(* IEC 61131-3 sources: Industry-PLC-LLM/data/PLCBEAD_repo/PLCBEAD_PLCEmbed-main/PLC-BEAD/Source/PLC_Programs (part 12) *)

(* ---- TEMP_EXT.ST ---- *)
FUNCTION UDINT_TO_TIME2:TIME

	VAR_INPUT
		IN :	UDINT;
	END_VAR

	UDINT_TO_TIME2 := DINT_TO_TIME(UDINT_TO_DINT(IN));

END_FUNCTION

FUNCTION_BLOCK T_PLC_MS_block
	VAR_OUTPUT
		T_PLC_MS :	UDINT;
	END_VAR

	VAR_EXTERNAL
		PLC_TICKS_PER_SEC :	INT;
		PLC_SYS_TICK_CNT :	DINT;
	END_VAR

	VAR
		debug :	BOOL;(*Debug-Mode ON / OFF*)
		N :	INT;(*Debug-Faktor*)
		Offset :	UDINT;(*Debug-Offset*)
		temp :	DWORD := DWORD#1;(*Debug-Offset*)
		mode :	BOOL;(*modus*)
		faktor :	UDINT;(*Systemtakt-Faktor*)
		init :	BOOL;
		v_plc_ticks_per_sec :	UDINT;
		base :	UDINT := UDINT#1000;
	END_VAR

	IF init = FALSE THEN
		v_plc_ticks_per_sec := INT_TO_UDINT(PLC_TICKS_PER_SEC);
		IF v_plc_ticks_per_sec = UDINT#1024 THEN
			faktor := UDINT#1;
			mode := FALSE;
		ELSIF v_plc_ticks_per_sec > UDINT#0 THEN
			IF v_plc_ticks_per_sec <= base THEN
				faktor := base / v_plc_ticks_per_sec;
				mode := FALSE;
			ELSE
				faktor := v_plc_ticks_per_sec / base;
				mode := TRUE;
			END_IF;
		ELSE
			faktor := UDINT#1;
		END_IF;
		init := TRUE;
	END_IF;

	IF mode THEN
		T_PLC_MS := DINT_TO_UDINT(PLC_SYS_TICK_CNT) / faktor;
	ELSE
		T_PLC_MS := DINT_TO_UDINT(PLC_SYS_TICK_CNT) * faktor;
	END_IF;

	IF debug THEN
		T_PLC_MS := (DWORD_TO_UDINT(SHL(UDINT_TO_DWORD(T_PLC_MS),N) OR SHL(temp,N)) - UDINT#1) + Offset;
	END_IF;
END_FUNCTION_BLOCK

FUNCTION _INT_TO_UDINT:UDINT
	VAR_INPUT
		IN :	INT;
	END_VAR

	_INT_TO_UDINT := DINT_TO_UDINT(INT_TO_DINT(IN));
END_FUNCTION

FUNCTION SET_DATE:UDINT

	VAR_INPUT
		YEAR :	INT;
		MONTH :	INT;
		DAY :	INT;
	END_VAR

	VAR
		count :	INT;
	END_VAR

	IF month > 2 THEN
		count := (month - 1) * 30;
		IF month > 7 THEN
			count := count + DWORD_TO_INT(SHR(DINT_TO_DWORD(INT_TO_DINT(month) - INT_TO_DINT(3)),1));
		ELSE
			count := count + DWORD_TO_INT(SHR(DINT_TO_DWORD(INT_TO_DINT(month) - INT_TO_DINT(4)),1));
		END_IF;
		IF SHL(INT_TO_WORD(year),14) = WORD#0 THEN
			count := count + 1;
		END_IF;
	ELSE
		count := (month - 1) * 31;
	END_IF;
	SET_DATE := (_INT_TO_UDINT(count + day - 1) + DWORD_TO_UDINT(SHR(UDINT_TO_DWORD(_INT_TO_UDINT(year) * UDINT#1461 - UDINT#2878169), 2))) * UDINT#86400;

END_FUNCTION

FUNCTION LEAP_OF_DATE:BOOL

	VAR_INPUT
		IDATE :	UDINT;
	END_VAR

	LEAP_OF_DATE := SHL(UDINT_TO_DWORD((idate + UDINT#43200) / UDINT#31557600), 30) = DWORD#16#80000000;

END_FUNCTION

FUNCTION DAY_OF_YEAR:INT
	VAR_INPUT
		IDATE :	DATE;
	END_VAR

	DAY_OF_YEAR := UDINT_TO_INT((DATE_TO_UDINT(idate) / UDINT#86400) MOD UDINT#1461);
	IF DAY_OF_YEAR > 729 THEN
		IF DAY_OF_YEAR > 1095 THEN DAY_OF_YEAR := DAY_OF_YEAR - 1095; ELSE DAY_OF_YEAR := DAY_OF_YEAR - 729; END_IF;
	ELSIF DAY_OF_YEAR > 364 THEN
		DAY_OF_YEAR := DAY_OF_YEAR - 364;
	ELSE
		DAY_OF_YEAR := DAY_OF_YEAR + 1;
	END_IF;
END_FUNCTION

FUNCTION DAY_OF_YEAR_UDINT:INT
	VAR_INPUT
		IDATE :	UDINT;
	END_VAR

	DAY_OF_YEAR_UDINT := UDINT_TO_INT((idate / UDINT#86400) MOD UDINT#1461);
	IF DAY_OF_YEAR_UDINT > 729 THEN
		IF DAY_OF_YEAR_UDINT > 1095 THEN DAY_OF_YEAR_UDINT := DAY_OF_YEAR_UDINT - 1095; ELSE DAY_OF_YEAR_UDINT := DAY_OF_YEAR_UDINT - 729; END_IF;
	ELSIF DAY_OF_YEAR_UDINT > 364 THEN
		DAY_OF_YEAR_UDINT := DAY_OF_YEAR_UDINT - 364;
	ELSE
		DAY_OF_YEAR_UDINT := DAY_OF_YEAR_UDINT + 1;
	END_IF;
END_FUNCTION

FUNCTION MONTH_OF_DATE_UDINT:INT

	VAR_INPUT
		IDATE :	UDINT;
	END_VAR

	MONTH_OF_DATE_UDINT := DAY_OF_YEAR_UDINT(idate);
	IF MONTH_OF_DATE_UDINT < 32 THEN
		MONTH_OF_DATE_UDINT := 1;
	ELSIF LEAP_OF_DATE(IDATE) THEN
		MONTH_OF_DATE_UDINT := (MONTH_OF_DATE_UDINT * 53 + 1668) / 1623;
	ELSE
		MONTH_OF_DATE_UDINT := (MONTH_OF_DATE_UDINT * 53 + 1700) / 1620;
	END_IF;

END_FUNCTION

FUNCTION DAY_OF_MONTH:INT
	VAR_INPUT
		IDATE :	UDINT;
	END_VAR

	day_of_month := day_of_year_UDINT(idate);

	IF leap_of_Date(idate) THEN
		CASE day_of_month OF
			32..60	:	day_of_month := day_of_month - 31;
			61..91	:	day_of_month := day_of_month - 60;
			92..121 :	day_of_month := day_of_month - 91;
			122..152:	day_of_month := day_of_month - 121;
			153..182:	day_of_month := day_of_month - 152;
			183..213:	day_of_month := day_of_month - 182;
			214..244:	day_of_month := day_of_month - 213;
			245..274:	day_of_month := day_of_month - 244;
			275..305:	day_of_month := day_of_month - 274;
			306..335:	day_of_month := day_of_month - 305;
			336..366:	day_of_month := day_of_month - 335;
		END_CASE;
	ELSE
		CASE day_of_month OF
			32..59	:	day_of_month := day_of_month - 31;
			60..90	:	day_of_month := day_of_month - 59;
			91..120 :	day_of_month := day_of_month - 90;
			121..151:	day_of_month := day_of_month - 120;
			152..181:	day_of_month := day_of_month - 151;
			182..212:	day_of_month := day_of_month - 181;
			213..243:	day_of_month := day_of_month - 212;
			244..273:	day_of_month := day_of_month - 243;
			274..304:	day_of_month := day_of_month - 273;
			305..334:	day_of_month := day_of_month - 304;
			335..365:	day_of_month := day_of_month - 334;
		END_CASE;
	END_IF;

END_FUNCTION

FUNCTION MID3:REAL

	VAR_INPUT
		IN1 :	REAL;
		IN2 :	REAL;
		IN3 :	REAL;
	END_VAR

	VAR
		_IN1 :	REAL;
		_IN2 :	REAL;
		_IN3 :	REAL;
	END_VAR

	_IN1 := IN1;
	_IN2 := IN2;
	_IN3 := IN3;

	IF _IN1 > _IN2 THEN MID3 := _IN1; _IN1 := _IN2; _IN2 := MID3; END_IF;
	IF _IN2 > _IN3 THEN _IN2 := _IN3; END_IF;
	MID3 := SEL(_IN1 > _IN2, _IN2, _IN1);

END_FUNCTION

FUNCTION _BYTE_TO_INT:INT
	VAR_INPUT
		IN :	BYTE;
	END_VAR

	_BYTE_TO_INT := USINT_TO_INT(BYTE_TO_USINT(IN));
END_FUNCTION

FUNCTION MULTI_IN:REAL

	VAR_INPUT
		IN_1 :	REAL;
		IN_2 :	REAL;
		IN_3 :	REAL;
		DEFAULT :	REAL;
		IN_MIN :	REAL;
		IN_MAX :	REAL;
		MODE :	BYTE;
	END_VAR

	VAR
		count :	INT;
		F1 :	BOOL;
		F2 :	BOOL;
		F3 :	BOOL;
	END_VAR

	F1 :=  in_1 > in_min AND in_1 < in_max;
	F2 :=  in_2 > in_min AND in_2 < in_max;
	F3 :=  in_3 > in_min AND in_3 < in_max;

	CASE _BYTE_TO_INT(mode) OF
	0:	count := 0;
		IF F1 THEN
			count := count + 1;
			MULTI_IN := in_1;
		ELSE
			MULTI_IN := 0.0;
		END_IF;
		IF F2 THEN
			count := count + 1;
			MULTI_IN := MULTI_IN + in_2;
		END_IF;
		IF F3 THEN
			count := count + 1;
			MULTI_IN := MULTI_IN + in_3;
		END_IF;
		MULTI_IN := SEL_REAL(count = 0, MULTI_IN / INT_TO_REAL(count), default);

	1:	MULTI_IN := SEL_REAL(F1, default, IN_1);

	2:	MULTI_IN := SEL_REAL(F2, default, IN_2);

	3:	MULTI_IN := SEL_REAL(F3, default, IN_3);

	4:	MULTI_IN := default;

	5:	MULTI_IN := SEL_REAL(F1, in_max, IN_1);
		IF F2 AND in_2 < MULTI_IN THEN MULTI_IN := in_2; END_IF;
		IF F3 AND in_3 < MULTI_IN THEN MULTI_IN := in_3; END_IF;
		IF MULTI_IN = in_max THEN MULTI_IN := default; END_IF;

	6:	MULTI_IN := SEL_REAL(F1, in_min, IN_1);
		IF F2 AND in_2 > MULTI_IN THEN MULTI_IN := in_2; END_IF;
		IF F3 AND in_3 > MULTI_IN THEN MULTI_IN := in_3; END_IF;
		IF MULTI_IN = in_min THEN MULTI_IN := default; END_IF;

	7:	IF F1 AND F2 AND F3 THEN MULTI_IN := MID3(in_1, in_2, in_3);
		ELSIF F1 AND F2 THEN MULTI_IN := MIN(in_1, in_2);
		ELSIF F1 AND F3 THEN MULTI_IN := MIN(in_1, in_3);
		ELSIF F2 AND F3 THEN MULTI_IN := MIN(in_2, in_3);
		ELSIF F1 THEN MULTI_IN := in_1;
		ELSIF F2 THEN MULTI_IN := in_2;
		ELSIF F3 THEN MULTI_IN := in_3;
		ELSE MULTI_IN := default;
		END_IF;

	END_CASE;

END_FUNCTION

FUNCTION _DT_TO_DATE_B:UDINT

	VAR_INPUT
		_INN :	UDINT;
	END_VAR

	_DT_TO_DATE_B := (_INN / UDINT#86400) * UDINT#86400;
END_FUNCTION

FUNCTION DT_TO_TOD2:UDINT
	VAR_INPUT
		IN :	UDINT;
	END_VAR

	DT_TO_TOD2 := (IN MOD UDINT#86400) * UDINT#1000;
END_FUNCTION

FUNCTION_BLOCK TEMP_EXT_Block

	VAR_INPUT
		T_EXT1 :	REAL;
		T_EXT2 :	REAL;
		T_EXT3 :	REAL;
		T_EXT_CONFIG :	BYTE := 0;
		DT_IN :	UDINT;
		T_EXT_MIN :	REAL := REAL#-40.0;
		T_EXT_MAX :	REAL := REAL#60.0;
		T_EXT_DEFAULT :	REAL := REAL#-10.0;
		HEAT_PERIOD_START :	UDINT := UDINT#20995200;
		HEAT_PERIOD_STOP :	UDINT := UDINT#10281600;
		COOL_PERIOD_START :	UDINT := UDINT#07776000;
		COOL_PERIOD_STOP :	UDINT := UDINT#23500800;
		HEAT_START_TEMP_DAY :	REAL := REAL#15.0;
		HEAT_START_TEMP_NIGHT :	REAL := REAL#10.0;
		HEAT_STOP_TEMP :	REAL := REAL#18.0;
		COOL_START_TEMP_DAY :	REAL := REAL#26.0;
		COOL_START_TEMP_NIGHT :	REAL := REAL#26.0;
		COOL_STOP_TEMP :	REAL := REAL#24.0;
		START_DAY :	UDINT := UDINT#32400000;
		START_NIGHT :	UDINT := UDINT#75600000;
		CYCLE_TIME :	TIME := t#10m;
	END_VAR

	VAR_OUTPUT
		T_EXT :	REAL;
		HEAT :	BOOL;
		COOL :	BOOL;
	END_VAR

	VAR
		tx :	TIME;
		last_run :	TIME;
		init :	BOOL;
		cool_start :	UDINT;
		cool_stop :	UDINT;
		heat_start :	UDINT;
		heat_stop :	UDINT;
		xdate :	UDINT;
		day :	BOOL;
		T_PLC_MS :	T_PLC_MS_Block;
	END_VAR

	IF NOT init THEN
		init := TRUE;
		heat_start := SET_DATE(1972,MONTH_OF_DATE_UDINT(heat_period_start),DAY_OF_MONTH(heat_period_start));
		heat_stop := SET_DATE(1972,MONTH_OF_DATE_UDINT(heat_period_stop),DAY_OF_MONTH(heat_period_stop));
		cool_start := SET_DATE(1972,MONTH_OF_DATE_UDINT(cool_period_start),DAY_OF_MONTH(cool_period_start));
		cool_stop := SET_DATE(1972,MONTH_OF_DATE_UDINT(cool_period_stop),DAY_OF_MONTH(cool_period_stop));
	END_IF;

	T_PLC_MS();
	tx:= UDINT_TO_TIME(T_PLC_MS.T_PLC_MS);

	IF tx - last_run < cycle_time THEN RETURN; END_IF;

	xdate := SET_DATE(1972,MONTH_OF_DATE_UDINT(_DT_TO_DATE_B(dt_in)),DAY_OF_MONTH(_DT_TO_DATE_B(dt_in)));
	day := DT_TO_TOD2(dt_in) >= start_day AND  DT_TO_TOD2(dt_in) < start_night;

	t_ext := MULTI_IN(t_ext1, t_ext2, t_ext3, t_ext_default, t_ext_min, t_ext_max, t_ext_config);

	IF (heat_start <= heat_stop AND xdate >= heat_start AND xdate <= heat_stop) OR (heat_start > heat_stop AND (xdate >= heat_start OR xdate <= heat_stop)) THEN
		IF day AND t_ext <= heat_start_temp_day THEN
			heat := TRUE;
		ELSIF NOT day AND t_ext <= heat_start_temp_night THEN
			heat := TRUE;
		ELSIF t_ext >= heat_stop_temp THEN
			heat := FALSE;
		END_IF;
	ELSE
		heat := FALSE;
	END_IF;

	IF (cool_start <= cool_stop AND xdate >= cool_start AND xdate <= cool_stop) OR (cool_start > cool_stop AND (xdate >= cool_start OR xdate <= cool_stop)) THEN
		IF day AND t_ext >= cool_start_temp_day THEN
			cool := TRUE;
		ELSIF NOT day AND t_ext >= cool_start_temp_night THEN
			cool := TRUE;
		ELSIF t_ext <= cool_stop_temp THEN
			cool := FALSE;
		END_IF;
	ELSE
		cool := FALSE;
	END_IF;

	last_run := tx;

END_FUNCTION_BLOCK

PROGRAM program0
	VAR
		T_EXT1 :	REAL;
		T_EXT2 :	REAL;
		T_EXT3 :	REAL;
		T_EXT_CONFIG :	BYTE := 0;
		DT_IN :	UDINT;
		T_EXT_MIN :	REAL := REAL#-40.0;
		T_EXT_MAX :	REAL := REAL#60.0;
		T_EXT_DEFAULT :	REAL := REAL#-10.0;
		HEAT_PERIOD_START :	UDINT := UDINT#20995200;
		HEAT_PERIOD_STOP :	UDINT := UDINT#10281600;
		COOL_PERIOD_START :	UDINT := UDINT#07776000;
		COOL_PERIOD_STOP :	UDINT := UDINT#23500800;
		HEAT_START_TEMP_DAY :	REAL := REAL#15.0;
		HEAT_START_TEMP_NIGHT :	REAL := REAL#10.0;
		HEAT_STOP_TEMP :	REAL := REAL#18.0;
		COOL_START_TEMP_DAY :	REAL := REAL#26.0;
		COOL_START_TEMP_NIGHT :	REAL := REAL#26.0;
		COOL_STOP_TEMP :	REAL := REAL#24.0;
		START_DAY :	UDINT := UDINT#32400000;
		START_NIGHT :	UDINT := UDINT#75600000;
		CYCLE_TIME :	TIME := t#10m;
		T_EXT :	REAL;
		HEAT :	BOOL;
		COOL :	BOOL;

		func_block : TEMP_EXT_Block;
	END_VAR

	func_block.T_EXT1 := T_EXT1;
	func_block.T_EXT2 := T_EXT2;
	func_block.T_EXT3 := T_EXT3 ;
	func_block.T_EXT_CONFIG := T_EXT_CONFIG;
	func_block.DT_IN := DT_IN;
	func_block.T_EXT_MIN := T_EXT_MIN ;
	func_block.T_EXT_MAX := T_EXT_MAX;
	func_block.T_EXT_DEFAULT := T_EXT_DEFAULT;
	func_block.HEAT_PERIOD_START := HEAT_PERIOD_START ;
	func_block.HEAT_PERIOD_STOP := HEAT_PERIOD_STOP;
	func_block.COOL_PERIOD_START := COOL_PERIOD_START;
	func_block.COOL_PERIOD_STOP := COOL_PERIOD_STOP ;
	func_block.HEAT_START_TEMP_DAY := HEAT_START_TEMP_DAY;
	func_block.HEAT_START_TEMP_NIGHT := HEAT_START_TEMP_NIGHT;
	func_block.HEAT_STOP_TEMP := HEAT_STOP_TEMP ;
	func_block.COOL_START_TEMP_DAY := COOL_START_TEMP_DAY;
	func_block.COOL_START_TEMP_NIGHT := COOL_START_TEMP_NIGHT;
	func_block.COOL_STOP_TEMP:= COOL_STOP_TEMP ;
	func_block.START_DAY := START_DAY;
	func_block.START_NIGHT := START_NIGHT;
	func_block.CYCLE_TIME:= CYCLE_TIME ;

	func_block();
	T_EXT  := func_block.T_EXT;
	HEAT  := func_block.HEAT;
	COOL  := func_block.COOL;

END_PROGRAM

CONFIGURATION Config0
	VAR_GLOBAL
		PLC_TICKS_PER_SEC :	INT;
		PLC_SYS_TICK_CNT :	DINT;
	END_VAR
  	RESOURCE Res0 ON PLC
    	TASK task0(INTERVAL := T#20ms,PRIORITY := 0);
    	PROGRAM instance0 WITH task0 : program0;
  	END_RESOURCE
END_CONFIGURATION

(* ---- TEMPERATURE.ST ---- *)
FUNCTION_BLOCK TEMPERATURE

	VAR_INPUT
		K :	REAL;
		C :	REAL := -273.15;
		F :	REAL := -459.67;
		RE :	REAL := -218.52;
		RA :	REAL := 0.0;
	END_VAR

	VAR_OUTPUT
		YK :	REAL;
		YC :	REAL;
		YF :	REAL;
		YRE :	REAL;
		YRA :	REAL;
	END_VAR

	YK := K + (C + 273.15) + (F + 459.67) * 0.555555555555 + (Re * 1.25 + 273.15) + (Ra * 0.555555555555);
	YC := YK -273.15;
	YF := YK * 1.8 - 459.67;
	YRe := (YK - 273.15) * 0.8;
	YRa := YK * 1.8;

END_FUNCTION_BLOCK

PROGRAM program0
  VAR
	K :	REAL;
	C :	REAL := -273.15;
	F :	REAL := -459.67;
	RE :	REAL := -218.52;
	RA :	REAL := 0.0;
	YK :	REAL;
	YC :	REAL;
	YF :	REAL;
	YRE :	REAL;
	YRA :	REAL;
	func_block : TEMPERATURE;
  END_VAR
	func_block.K  :=K;
	func_block.C  :=C;
	func_block.F  :=F;
	func_block.RE  :=RE;
	func_block.RA  :=RA;
	func_block();
	YK := func_block.YK;
	YC := func_block.YC;
	YF := func_block.YF;
	YRE := func_block.YRE;
	YRA := func_block.YRA;

END_PROGRAM

CONFIGURATION Config0
	RESOURCE Res0 ON PLC
		TASK task0(INTERVAL := T#20ms,PRIORITY := 0);
		PROGRAM instance0 WITH task0 : program0;
	END_RESOURCE
END_CONFIGURATION

(* ---- TICKER.ST ---- *)
TYPE
	oscat_delay_buf             : ARRAY [0..31]   OF REAL;
END_TYPE

FUNCTION INC1:INT

	VAR_INPUT
		X :	INT;
		N :	INT;
	END_VAR

	IF X >= N - 1 THEN
		INC1 := 0;
	ELSE
		INC1 := X + 1;
	END_IF;
END_FUNCTION

FUNCTION_BLOCK DELAY

	VAR_INPUT
		IN :	REAL;
		N :	INT;
		RST :	BOOL;
	END_VAR

	VAR_OUTPUT
		OUT :	REAL;
	END_VAR

	VAR
		buf :	oscat_delay_buf;
		i :	INT;
		init :	BOOL;
		stop :	INT;
	END_VAR

	stop := LIMIT(0,N,32) - 1;
	IF rst OR NOT init THEN
		init := TRUE;
		FOR i := 0 TO stop DO buf[i] := in; END_FOR;
		out := in;
		i := 0;
	ELSIF stop < 0 THEN
		out := in;
	ELSE
		out := buf[i];
		buf[i] := in;
		i := INC1(i, N);
	END_IF;

END_FUNCTION_BLOCK

FUNCTION_BLOCK TICKER

	VAR_INPUT
		N :	INT;
		PT :	TIME;
		TEXT :	STRING;
	END_VAR

	VAR_OUTPUT
		DISPLAY :	STRING;
	END_VAR

	VAR
		_delay :	TP;
		rollout :	STRING;
		text_len :	INT;
		rollout_step :	INT;
		_step :	INT;
	END_VAR

	text_len := LEN(text);

	IF N < text_len THEN
		IF NOT _delay.Q THEN

			IF _step > text_len THEN
				rollout_step := 0;
				rollout := '';
				_step := 0;
			END_IF;

			IF _step + N > text_len THEN
				_step := _step + 1;
				rollout_step := rollout_step +1;
				display := MID(text, N - rollout_step, _step);
				rollout := CONCAT(rollout,'#');
				display := CONCAT(display,rollout);
			ELSE
				_step := _step + 1;
				display := MID(text, N, _step);
			END_IF;
			_delay(TRUE, PT);
		ELSE
			_delay(FALSE);
		END_IF;
	ELSE
		display := text;
	END_IF;

END_FUNCTION_BLOCK

PROGRAM program0
	VAR
		N :	INT;
		PT :	TIME;
		TEXT :	STRING;
		DISPLAY :	STRING;
		func_block : TICKER;
  	END_VAR
	func_block.N  :=N;
	func_block.PT  :=PT;
	func_block.TEXT  :=TEXT;
	func_block();
	DISPLAY := func_block.DISPLAY;
END_PROGRAM

CONFIGURATION Config0
	RESOURCE Res0 ON PLC
		TASK task0(INTERVAL := T#20ms,PRIORITY := 0);
		PROGRAM instance0 WITH task0 : program0;
	END_RESOURCE
END_CONFIGURATION

(* ---- TIMER_1.ST ---- *)
FUNCTION TIMECHECK:BOOL

	VAR_INPUT
		TD :	UDINT;
		START :	UDINT;
		STOP :	UDINT;
	END_VAR

	IF stop < start THEN
		TIMECHECK := start <= TD OR  TD < stop;
	ELSE
		TIMECHECK := start <= TD AND TD < stop;
	END_IF;

END_FUNCTION

FUNCTION TIME_TO_TOD:UDINT

	VAR_INPUT
		IN :	TIME;
	END_VAR

	TIME_TO_TOD := DWORD_TO_UDINT(TIME_TO_DWORD(IN));
END_FUNCTION

FUNCTION TOD_TO_TIME:TIME
	VAR_INPUT
		IN :	UDINT;
	END_VAR

	TOD_TO_TIME := DWORD_TO_TIME(UDINT_TO_DWORD(IN));
END_FUNCTION

FUNCTION DAY_OF_WEEK:INT
  VAR_INPUT
    IDATE :	UDINT;
  END_VAR

  DAY_OF_WEEK := UDINT_TO_INT((idate / UDINT#86400 + UDINT#3) MOD UDINT#7) + INT#01;
END_FUNCTION

FUNCTION _DT_TO_DATE_B:UDINT

	VAR_INPUT
		_INN :	UDINT;
	END_VAR

	_DT_TO_DATE_B := (_INN / UDINT#86400) * UDINT#86400;
END_FUNCTION

FUNCTION DT_TO_TOD2:UDINT
	VAR_INPUT
		IN :	UDINT;
	END_VAR

	DT_TO_TOD2 := (IN MOD UDINT#86400) * UDINT#1000;
END_FUNCTION

FUNCTION TIME_TO_TOD2:UDINT

	VAR_INPUT
		IN :	TIME;
	END_VAR

	TIME_TO_TOD2 := DWORD_TO_UDINT(TIME_TO_DWORD(IN));
END_FUNCTION

FUNCTION_BLOCK TIMER_1_Block

	VAR_INPUT
		E :	BOOL := TRUE;
		DTI :	UDINT;
		START :	UDINT;
		DURATION :	TIME;
		DAY :	BYTE := BYTE#2#0111_1111;
	END_VAR

	VAR_OUTPUT
		Q :	BOOL;
		STOP :	TIME;
	END_VAR

	IF E THEN
		stop := TOD_TO_TIME(START) + DURATION;
		IF stop > T#24h THEN stop := stop - T#24h; END_IF;
		Q := TIMECHECK(DT_TO_TOD2(DTI), START, TIME_TO_TOD2(stop)) AND (SHR(BYTE#128, DAY_OF_WEEK(_DT_TO_DATE_B(DTI))) AND DAY) > BYTE#0;
	ELSE
		Q := FALSE;
	END_IF;

END_FUNCTION_BLOCK

PROGRAM program0
	VAR
		E :	BOOL := TRUE;
		DTI :	UDINT;
		START :	UDINT;
		DURATION :	TIME;
		DAY :	BYTE := BYTE#2#0111_1111;
		Q :	BOOL;
		STOP :	TIME;

		func_block : TIMER_1_Block;
	END_VAR
	func_block.E := E;
	func_block.DTI := DTI;
	func_block.START := START ;
	func_block.DURATION    := DURATION    ;
	func_block.DAY := DAY;

	func_block();
	Q  := func_block.Q;
	STOP  := func_block.STOP;
END_PROGRAM

CONFIGURATION Config0
	RESOURCE Res0 ON PLC
		TASK task0(INTERVAL := T#20ms,PRIORITY := 0);
		PROGRAM instance0 WITH task0 : program0;
	END_RESOURCE
END_CONFIGURATION

(* ---- TIMER_2.ST ---- *)
FUNCTION UDINT_TO_TIME2:TIME

	VAR_INPUT
		IN :	UDINT;
	END_VAR

	UDINT_TO_TIME2 := DINT_TO_TIME(UDINT_TO_DINT(IN));

END_FUNCTION

FUNCTION_BLOCK T_PLC_MS_block
	VAR_OUTPUT
		T_PLC_MS :	UDINT;
	END_VAR

	VAR_EXTERNAL
		PLC_TICKS_PER_SEC :	INT;
		PLC_SYS_TICK_CNT :	DINT;
	END_VAR

	VAR
		debug :	BOOL;(*Debug-Mode ON / OFF*)
		N :	INT;(*Debug-Faktor*)
		Offset :	UDINT;(*Debug-Offset*)
		temp :	DWORD := DWORD#1;(*Debug-Offset*)
		mode :	BOOL;(*modus*)
		faktor :	UDINT;(*Systemtakt-Faktor*)
		init :	BOOL;
		v_plc_ticks_per_sec :	UDINT;
		base :	UDINT := UDINT#1000;
	END_VAR

	IF init = FALSE THEN
		v_plc_ticks_per_sec := INT_TO_UDINT(PLC_TICKS_PER_SEC);
		IF v_plc_ticks_per_sec = UDINT#1024 THEN
			faktor := UDINT#1;
			mode := FALSE;
		ELSIF v_plc_ticks_per_sec > UDINT#0 THEN
			IF v_plc_ticks_per_sec <= base THEN
				faktor := base / v_plc_ticks_per_sec;
				mode := FALSE;
			ELSE
				faktor := v_plc_ticks_per_sec / base;
				mode := TRUE;
			END_IF;
		ELSE
			faktor := UDINT#1;
		END_IF;
		init := TRUE;
	END_IF;

	IF mode THEN
		T_PLC_MS := DINT_TO_UDINT(PLC_SYS_TICK_CNT) / faktor;
	ELSE
		T_PLC_MS := DINT_TO_UDINT(PLC_SYS_TICK_CNT) * faktor;
	END_IF;

	IF debug THEN
		T_PLC_MS := (DWORD_TO_UDINT(SHL(UDINT_TO_DWORD(T_PLC_MS),N) OR SHL(temp,N)) - UDINT#1) + Offset;
	END_IF;
END_FUNCTION_BLOCK

FUNCTION DAY_OF_WEEK:INT
  VAR_INPUT
    IDATE :	UDINT;
  END_VAR

  DAY_OF_WEEK := UDINT_TO_INT((idate / UDINT#86400 + UDINT#3) MOD UDINT#7) + INT#01;
END_FUNCTION

FUNCTION _BYTE_TO_INT:INT
	VAR_INPUT
		IN :	BYTE;
	END_VAR

	_BYTE_TO_INT := USINT_TO_INT(BYTE_TO_USINT(IN));
END_FUNCTION

FUNCTION LEAP_OF_DATE:BOOL

	VAR_INPUT
		IDATE :	UDINT;
	END_VAR

	LEAP_OF_DATE := SHL(UDINT_TO_DWORD((idate + UDINT#43200) / UDINT#31557600), 30) = DWORD#16#80000000;

END_FUNCTION

FUNCTION DAY_OF_YEAR:INT
	VAR_INPUT
		IDATE :	DATE;
	END_VAR

	DAY_OF_YEAR := UDINT_TO_INT((DATE_TO_UDINT(idate) / UDINT#86400) MOD UDINT#1461);
	IF DAY_OF_YEAR > 729 THEN
		IF DAY_OF_YEAR > 1095 THEN DAY_OF_YEAR := DAY_OF_YEAR - 1095; ELSE DAY_OF_YEAR := DAY_OF_YEAR - 729; END_IF;
	ELSIF DAY_OF_YEAR > 364 THEN
		DAY_OF_YEAR := DAY_OF_YEAR - 364;
	ELSE
		DAY_OF_YEAR := DAY_OF_YEAR + 1;
	END_IF;
END_FUNCTION

FUNCTION DAY_OF_YEAR_UDINT:INT
	VAR_INPUT
		IDATE :	UDINT;
	END_VAR

	DAY_OF_YEAR_UDINT := UDINT_TO_INT((idate / UDINT#86400) MOD UDINT#1461);
	IF DAY_OF_YEAR_UDINT > 729 THEN
		IF DAY_OF_YEAR_UDINT > 1095 THEN DAY_OF_YEAR_UDINT := DAY_OF_YEAR_UDINT - 1095; ELSE DAY_OF_YEAR_UDINT := DAY_OF_YEAR_UDINT - 729; END_IF;
	ELSIF DAY_OF_YEAR_UDINT > 364 THEN
		DAY_OF_YEAR_UDINT := DAY_OF_YEAR_UDINT - 364;
	ELSE
		DAY_OF_YEAR_UDINT := DAY_OF_YEAR_UDINT + 1;
	END_IF;
END_FUNCTION

FUNCTION MONTH_OF_DATE_UDINT:INT

	VAR_INPUT
		IDATE :	UDINT;
	END_VAR

	MONTH_OF_DATE_UDINT := DAY_OF_YEAR_UDINT(idate);
	IF MONTH_OF_DATE_UDINT < 32 THEN
		MONTH_OF_DATE_UDINT := 1;
	ELSIF LEAP_OF_DATE(IDATE) THEN
		MONTH_OF_DATE_UDINT := (MONTH_OF_DATE_UDINT * 53 + 1668) / 1623;
	ELSE
		MONTH_OF_DATE_UDINT := (MONTH_OF_DATE_UDINT * 53 + 1700) / 1620;
	END_IF;

END_FUNCTION

FUNCTION DAY_OF_MONTH:INT
	VAR_INPUT
		IDATE :	UDINT;
	END_VAR

	day_of_month := day_of_year_UDINT(idate);

	IF leap_of_Date(idate) THEN
		CASE day_of_month OF
			32..60	:	day_of_month := day_of_month - 31;
			61..91	:	day_of_month := day_of_month - 60;
			92..121 :	day_of_month := day_of_month - 91;
			122..152:	day_of_month := day_of_month - 121;
			153..182:	day_of_month := day_of_month - 152;
			183..213:	day_of_month := day_of_month - 182;
			214..244:	day_of_month := day_of_month - 213;
			245..274:	day_of_month := day_of_month - 244;
			275..305:	day_of_month := day_of_month - 274;
			306..335:	day_of_month := day_of_month - 305;
			336..366:	day_of_month := day_of_month - 335;
		END_CASE;
	ELSE
		CASE day_of_month OF
			32..59	:	day_of_month := day_of_month - 31;
			60..90	:	day_of_month := day_of_month - 59;
			91..120 :	day_of_month := day_of_month - 90;
			121..151:	day_of_month := day_of_month - 120;
			152..181:	day_of_month := day_of_month - 151;
			182..212:	day_of_month := day_of_month - 181;
			213..243:	day_of_month := day_of_month - 212;
			244..273:	day_of_month := day_of_month - 243;
			274..304:	day_of_month := day_of_month - 273;
			305..334:	day_of_month := day_of_month - 304;
			335..365:	day_of_month := day_of_month - 334;
		END_CASE;
	END_IF;

END_FUNCTION

FUNCTION MONTH_OF_DATE:INT

	VAR_INPUT
		IDATE :	DATE;
	END_VAR

	MONTH_OF_DATE := DAY_OF_YEAR(idate);
	IF MONTH_OF_DATE < 32 THEN
		MONTH_OF_DATE := 1;
	ELSIF LEAP_OF_DATE(DATE_TO_UDINT(IDATE)) THEN
		MONTH_OF_DATE := (MONTH_OF_DATE * 53 + 1668) / 1623;
	ELSE
		MONTH_OF_DATE := (MONTH_OF_DATE * 53 + 1700) / 1620;
	END_IF;

END_FUNCTION

FUNCTION TIME_TO_UDINT2:UDINT
	VAR_INPUT
		X :	TIME;
	END_VAR

	TIME_TO_UDINT2 := DINT_TO_UDINT(TIME_TO_DINT(X));
END_FUNCTION

FUNCTION DT_TO_TOD2:UDINT
	VAR_INPUT
		IN :	UDINT;
	END_VAR

	DT_TO_TOD2 := (IN MOD UDINT#86400) * UDINT#1000;
END_FUNCTION

FUNCTION _DT_TO_DATE_B:UDINT

	VAR_INPUT
		_INN :	UDINT;
	END_VAR

	_DT_TO_DATE_B := (_INN / UDINT#86400) * UDINT#86400;
END_FUNCTION

FUNCTION_BLOCK TIMER_2_Block

	VAR_INPUT
		DT_IN :	UDINT;
		START :	UDINT;
		DURATION :	TIME;
		MODE :	BYTE;
		HOLIDAY :	BOOL;
	END_VAR

	VAR_OUTPUT
		Q :	BOOL;
	END_VAR

	VAR
		last_check :	TIME := T#0s;
		dat :	UDINT;
		daytime :	UDINT;
		activation :	TIME;
		tx :	TIME;
		enabled :	BOOL;
		wday :	INT;
		init :	BOOL;
	END_VAR

	VAR RETAIN
		run_date :	UDINT;
	END_VAR

	VAR
		T_PLC_MS :	T_PLC_MS_Block;
	END_VAR

	T_PLC_MS();
	tx:= UDINT_TO_TIME(T_PLC_MS.T_PLC_MS);

	IF NOT init THEN
		init := TRUE;
		last_check := tx - t#100ms;
	END_IF;

	IF tx - last_check < T#100ms THEN RETURN; END_IF;

	dat := _DT_TO_DATE_B(dt_in);
	daytime := DT_TO_TOD2(dt_in);
	wday := DAY_OF_WEEK(dat);

	CASE _BYTE_TO_INT(mode) OF
	1..7:
		enabled := wday = _BYTE_TO_INT(mode);
	11:
		enabled := TRUE;
	12..16:
		enabled := (dat / UDINT#86400) MOD (BYTE_TO_UDINT(mode) - UDINT#10) = UDINT#0;
	20:
		enabled := wday <= 5;
	21:
		enabled := wday > 5;
	22:
		enabled := wday <= 5 AND NOT holiday;
	23:
		enabled := wday > 5 OR holiday;
	24:
		enabled := holiday;
	25:
		enabled := DAY_OF_MONTH(dat) = 1;
	26:
		enabled := day_of_month(dat + TIME_TO_UDINT2(t#1d)) = 1;
	27:
		enabled := DAY_OF_MONTH(dat) = 31 AND MONTH_OF_DATE_UDINT(dat) = 12;
	28:
		enabled := DAY_OF_YEAR_UDINT(dat) = 1;
	ELSE
		enabled := FALSE;
	END_CASE;

	IF enabled AND NOT Q AND daytime >= start AND run_date <> dat THEN
		Q := TRUE;
		activation := tx;
		run_date := dat;
	ELSIF Q AND tx - activation >= duration THEN
		Q := FALSE;
	END_IF;
	last_check := Tx;

END_FUNCTION_BLOCK

PROGRAM program0
	VAR
		DT_IN :	UDINT;
		START :	UDINT;
		DURATION :	TIME;
		MODE :	BYTE;
		HOLIDAY :	BOOL;
		Q :	BOOL;

		func_block : TIMER_2_Block;
	END_VAR
	func_block.DT_IN := DT_IN;
	func_block.START := START;
	func_block.DURATION := DURATION ;
	func_block.MODE    := MODE    ;
	func_block.HOLIDAY := HOLIDAY;

	func_block();
	Q  := func_block.Q;
END_PROGRAM

CONFIGURATION Config0
	VAR_GLOBAL
		PLC_TICKS_PER_SEC :	INT;
		PLC_SYS_TICK_CNT :	DINT;
	END_VAR
  	RESOURCE Res0 ON PLC
    	TASK task0(INTERVAL := T#20ms,PRIORITY := 0);
    	PROGRAM instance0 WITH task0 : program0;
  	END_RESOURCE
END_CONFIGURATION

(* ---- TIMER_EXT.ST ---- *)
FUNCTION_BLOCK MANUAL_2_Block

	VAR_INPUT
		_IN :	BOOL;
		ENA :	BOOL;
		_ON :	BOOL;
		OFF :	BOOL;
		MAN :	BOOL;
	END_VAR

	VAR_OUTPUT
		Q :	BOOL;
		STATUS :	BYTE;
	END_VAR

	IF ena THEN
		IF NOT _ON AND NOT OFF THEN
			Q := _IN;
			STATUS := BYTE#100;
		ELSIF _on AND NOT off THEN
			Q := TRUE;
			STATUS := BYTE#101;
		ELSIF NOT _on AND off THEN
			q := FALSE;
			STATUS := BYTE#102;
		ELSE
			Q := MAN;
			STATUS := BYTE#103;
		END_IF;
	ELSE
		Q := FALSE;
		STATUS := BYTE#104;
	END_IF;

END_FUNCTION_BLOCK

FUNCTION_BLOCK DEBOUNCE_Block

	VAR_INPUT
		IN :	BOOL;
		TD :	TIME;
		PM :	BOOL;
	END_VAR

	VAR_OUTPUT
		Q :	BOOL;
	END_VAR

	VAR
		deb :	TOF;
	END_VAR

	IF NOT deb.Q AND IN THEN
		Q := TRUE;
	ELSIF NOT PM THEN
		Q := deb.Q;
	ELSE
		Q := FALSE;
	END_IF;

END_FUNCTION_BLOCK

FUNCTION_BLOCK T_PLC_MS_block

	VAR_OUTPUT
		T_PLC_MS :	UDINT;
	END_VAR

	VAR_EXTERNAL
		PLC_TICKS_PER_SEC :	INT;
		PLC_SYS_TICK_CNT :	DINT;
	END_VAR

	VAR
		debug :	BOOL;(*Debug-Mode ON / OFF*)
		N :	INT;(*Debug-Faktor*)
		Offset :	UDINT;(*Debug-Offset*)
		temp :	DWORD := DWORD#1;(*Debug-Offset*)
		mode :	BOOL;(*modus*)
		faktor :	UDINT;(*Systemtakt-Faktor*)
		init :	BOOL;
		v_plc_ticks_per_sec :	UDINT;
		base :	UDINT := UDINT#1000;
	END_VAR

	IF init = FALSE THEN
		v_plc_ticks_per_sec := INT_TO_UDINT(PLC_TICKS_PER_SEC);
		IF v_plc_ticks_per_sec = UDINT#1024 THEN
			faktor := UDINT#1;
			mode := FALSE;
		ELSIF v_plc_ticks_per_sec > UDINT#0 THEN
			IF v_plc_ticks_per_sec <= base THEN
				faktor := base / v_plc_ticks_per_sec;
				mode := FALSE;
			ELSE
				faktor := v_plc_ticks_per_sec / base;
				mode := TRUE;
			END_IF;
		ELSE
			faktor := UDINT#1;
		END_IF;
		init := TRUE;
	END_IF;

	IF mode THEN
		T_PLC_MS := DINT_TO_UDINT(PLC_SYS_TICK_CNT) / faktor;
	ELSE
		T_PLC_MS := DINT_TO_UDINT(PLC_SYS_TICK_CNT) * faktor;
	END_IF;

	IF debug THEN
		T_PLC_MS := (DWORD_TO_UDINT(SHL(UDINT_TO_DWORD(T_PLC_MS),N) OR SHL(temp,N)) - UDINT#1) + Offset;
	END_IF;

END_FUNCTION_BLOCK

FUNCTION DT_TO_TOD2:UDINT
	VAR_INPUT
		IN :	UDINT;
	END_VAR

	DT_TO_TOD2 := (IN MOD UDINT#86400) * UDINT#1000;
END_FUNCTION

FUNCTION _DT_TO_DATE_B:UDINT

	VAR_INPUT
		_INN :	UDINT;
	END_VAR

	_DT_TO_DATE_B := (_INN / UDINT#86400) * UDINT#86400;
END_FUNCTION

FUNCTION DAY_OF_WEEK:INT
  VAR_INPUT
    IDATE :	UDINT;
  END_VAR

  DAY_OF_WEEK := UDINT_TO_INT((idate / UDINT#86400 + UDINT#3) MOD UDINT#7) + INT#01;
END_FUNCTION

FUNCTION TIME_TO_UDINT2:UDINT
	VAR_INPUT
		X :	TIME;
	END_VAR

	TIME_TO_UDINT2 := DINT_TO_UDINT(TIME_TO_DINT(X));
END_FUNCTION

FUNCTION_BLOCK TIMER_EXT_Block

	VAR_INPUT
		ENA :	BOOL;
		_ON :	BOOL;
		OFF :	BOOL;
		MAN :	BOOL;
		SWITCH :	BOOL;
		DT_IN :	UDINT;
		SUN_SET :	UDINT;
		SUN_RISE :	UDINT;
		HOLIDAY :	BOOL;
		T_DEBOUNCE :	TIME := T#100ms;
		T_RISE_START :	TIME;
		T_RISE_STOP :	TIME;
		T_SET_START :	TIME;
		T_SET_STOP :	TIME;
		T_DAY_START :	UDINT;
		T_DAY_STOP :	UDINT;
		ENABLE_SATURDAY :	BOOL;
		ENABLE_SUNDAY :	BOOL;
		ENABLE_HOLIDAY :	BOOL;
	END_VAR

	VAR_OUTPUT
		Q :	BOOL;
		STATUS :	BYTE;
	END_VAR

	VAR
		mx :	MANUAL_2_Block;
		deb :	DEBOUNCE_Block;
		tdx :	UDINT;
		wdx :	INT;
		tc :	TIME;
		tx :	UDINT;
		tl :	UDINT;
		qx :	BOOL;
		T_PLC_MS :	T_PLC_MS_Block;
		init :	BOOL;
	END_VAR

	SUN_RISE := SUN_RISE / UDINT#1000 * UDINT#1000;
	SUN_SET := SUN_SET / UDINT#1000 * UDINT#1000;

	T_PLC_MS();
	tx:= T_PLC_MS.T_PLC_MS;
	IF NOT init THEN
		init := TRUE;
		tl := tx;
	END_IF;
	tc := UDINT_TO_TIME(tx - tl);
	IF tc < t#200ms THEN RETURN; END_IF;
	tl := tx;

	deb(in := SWITCH, TD := T_DEBOUNCE, PM := TRUE);

	tdx := DT_TO_TOD2(dt_in);
	wdx := DAY_OF_WEEK(_DT_TO_DATE_B(dt_in));

	IF deb.Q THEN
		qx := NOT qx;
		status := BYTE#110;
	ELSIF holiday AND NOT enable_holiday THEN
		qx := FALSE;
	ELSIF wdx = 6 AND NOT enable_saturday THEN
		qx := FALSE;
	ELSIF wdx = 7 AND NOT enable_sunday THEN
		qx := FALSE;
	ELSIF T_day_start > UDINT#00 AND tdx - T_DAY_START <= TIME_TO_UDINT2(tc) THEN
		qx := TRUE;
		status := BYTE#111;
	ELSIF T_DAY_STOP > UDINT#00 AND tdx - T_DAY_STOP <= TIME_TO_UDINT2(tc) THEN
		qx := FALSE;
		status := BYTE#112;
	ELSIF T_RISE_START > T#0s AND tdx - SUN_RISE + TIME_TO_UDINT2(T_RISE_START) <= TIME_TO_UDINT2(tc) THEN
		qx := TRUE;
		status := BYTE#113;
	ELSIF T_RISE_STOP > T#0s AND tdx - SUN_RISE - TIME_TO_UDINT2(T_RISE_STOP) <= TIME_TO_UDINT2(tc) THEN
		qx := FALSE;
		status := BYTE#114;
	ELSIF T_SET_start > T#0s AND tdx - SUN_SET + TIME_TO_UDINT2(T_SET_START) <= TIME_TO_UDINT2(tc) THEN
		qx := TRUE;
		status := BYTE#115;
	ELSIF T_SET_STOP > T#0s AND tdx - SUN_SET - TIME_TO_UDINT2(T_SET_STOP) <= TIME_TO_UDINT2(tc) THEN
		qx := FALSE;
		status := BYTE#116;
	END_IF;

	mx(_IN := qx, ena := ENA, _ON := _ON, off := OFF, man := MAN);
	Q := mx.Q;

	IF mx.STATUS > BYTE#100 THEN status := mx.STATUS; END_IF;

END_FUNCTION_BLOCK

PROGRAM program0
	VAR
		ENA :	BOOL;
		_ON :	BOOL;
		OFF :	BOOL;
		MAN :	BOOL;
		SWITCH :	BOOL;
		DT_IN :	UDINT;
		SUN_SET :	UDINT;
		SUN_RISE :	UDINT;
		HOLIDAY :	BOOL;
		T_DEBOUNCE :	TIME := T#100ms;
		T_RISE_START :	TIME;
		T_RISE_STOP :	TIME;
		T_SET_START :	TIME;
		T_SET_STOP :	TIME;
		T_DAY_START :	UDINT;
		T_DAY_STOP :	UDINT;
		ENABLE_SATURDAY :	BOOL;
		ENABLE_SUNDAY :	BOOL;
		ENABLE_HOLIDAY :	BOOL;
		Q :	BOOL;
		STATUS :	BYTE;

		func_block : TIMER_EXT_Block;
	END_VAR
	func_block.ENA := ENA;
	func_block._ON := _ON;
	func_block.OFF := OFF ;
	func_block.MAN    := MAN    ;
	func_block.SWITCH := SWITCH;
	func_block.DT_IN := DT_IN;
	func_block.SUN_SET := SUN_SET;
	func_block.SUN_RISE := SUN_RISE ;
	func_block.HOLIDAY    := HOLIDAY    ;
	func_block.T_DEBOUNCE := T_DEBOUNCE;
	func_block.T_RISE_START := T_RISE_START;
	func_block.T_RISE_STOP := T_RISE_STOP;
	func_block.T_SET_START := T_SET_START ;
	func_block.T_SET_STOP    := T_SET_STOP    ;
	func_block.T_DAY_START := T_DAY_START;
	func_block.T_DAY_STOP := T_DAY_STOP;
	func_block.ENABLE_SATURDAY := ENABLE_SATURDAY;
	func_block.ENABLE_SUNDAY := ENABLE_SUNDAY ;
	func_block.ENABLE_HOLIDAY    := ENABLE_HOLIDAY    ;

	func_block();
	Q  := func_block.Q;
	STATUS := func_block.STATUS;
END_PROGRAM

CONFIGURATION Config0
	VAR_GLOBAL
		PLC_TICKS_PER_SEC :	INT;
		PLC_SYS_TICK_CNT :	DINT;
	END_VAR
  	RESOURCE Res0 ON PLC
    	TASK task0(INTERVAL := T#20ms,PRIORITY := 0);
    	PROGRAM instance0 WITH task0 : program0;
  	END_RESOURCE
END_CONFIGURATION

(* ---- TMAX.ST ---- *)
FUNCTION UDINT_TO_TIME2:TIME

	VAR_INPUT
		IN :	UDINT;
	END_VAR

	UDINT_TO_TIME2 := DINT_TO_TIME(UDINT_TO_DINT(IN));

END_FUNCTION

FUNCTION_BLOCK T_PLC_MS_block
	VAR_OUTPUT
		T_PLC_MS :	UDINT;
	END_VAR

	VAR_EXTERNAL
		PLC_TICKS_PER_SEC :	INT;
		PLC_SYS_TICK_CNT :	DINT;
	END_VAR

	VAR
		debug :	BOOL;(*Debug-Mode ON / OFF*)
		N :	INT;(*Debug-Faktor*)
		Offset :	UDINT;(*Debug-Offset*)
		temp :	DWORD := DWORD#1;(*Debug-Offset*)
		mode :	BOOL;(*modus*)
		faktor :	UDINT;(*Systemtakt-Faktor*)
		init :	BOOL;
		v_plc_ticks_per_sec :	UDINT;
		base :	UDINT := UDINT#1000;
	END_VAR

	IF init = FALSE THEN
		v_plc_ticks_per_sec := INT_TO_UDINT(PLC_TICKS_PER_SEC);
		IF v_plc_ticks_per_sec = UDINT#1024 THEN
			faktor := UDINT#1;
			mode := FALSE;
		ELSIF v_plc_ticks_per_sec > UDINT#0 THEN
			IF v_plc_ticks_per_sec <= base THEN
				faktor := base / v_plc_ticks_per_sec;
				mode := FALSE;
			ELSE
				faktor := v_plc_ticks_per_sec / base;
				mode := TRUE;
			END_IF;
		ELSE
			faktor := UDINT#1;
		END_IF;
		init := TRUE;
	END_IF;

	IF mode THEN
		T_PLC_MS := DINT_TO_UDINT(PLC_SYS_TICK_CNT) / faktor;
	ELSE
		T_PLC_MS := DINT_TO_UDINT(PLC_SYS_TICK_CNT) * faktor;
	END_IF;

	IF debug THEN
		T_PLC_MS := (DWORD_TO_UDINT(SHL(UDINT_TO_DWORD(T_PLC_MS),N) OR SHL(temp,N)) - UDINT#1) + Offset;
	END_IF;

END_FUNCTION_BLOCK

FUNCTION_BLOCK TMAX

	VAR_INPUT
		IN :	BOOL;
		PT :	TIME;
	END_VAR

	VAR_OUTPUT
		Q :	BOOL;
		Z :	BOOL;
	END_VAR

	VAR
		tx :	TIME;
		start :	TIME;
		last_in :	BOOL;
		T_PLC_MS :	T_PLC_MS_block;
	END_VAR

	T_PLC_MS();
	tx:= UDINT_TO_TIME(T_PLC_MS.T_PLC_MS);

	Z := FALSE;

	IF NOT in THEN
		Q := FALSE;
	ELSIF IN AND NOT last_in THEN
		Q := TRUE;
		start := tx;
	ELSIF (tx - start >= PT) AND Q THEN
		Q := FALSE;
		Z := TRUE;
	END_IF;

	last_in := IN;

END_FUNCTION_BLOCK

PROGRAM program0
  VAR
	IN :	BOOL;
	PT :	TIME;
	Q :	BOOL;
	Z :	BOOL;
	func_block : TMAX;
  END_VAR
	func_block.IN  :=IN;
	func_block.PT  :=PT;
	func_block();
	Q := func_block.Q;
	Z := func_block.Z;

END_PROGRAM

CONFIGURATION Config0
	VAR_GLOBAL
		PLC_TICKS_PER_SEC :	INT;
		PLC_SYS_TICK_CNT :	DINT;
	END_VAR
	RESOURCE Res0 ON PLC
		TASK task0(INTERVAL := T#20ms,PRIORITY := 0);
		PROGRAM instance0 WITH task0 : program0;
	END_RESOURCE
END_CONFIGURATION

(* ---- TMIN.ST ---- *)
FUNCTION_BLOCK TMIN

	VAR_INPUT
		IN :	BOOL;
		PT :	TIME;
	END_VAR

	VAR_OUTPUT
		Q :	BOOL;
	END_VAR

	VAR
		pm :	TP;
	END_VAR

	pm(in := IN, PT := PT);
	Q := IN OR pm.Q;

END_FUNCTION_BLOCK

PROGRAM program0
  VAR
	IN :	BOOL;
	PT :	TIME;
	Q :	BOOL;
	func_block : TMIN;
  END_VAR
	func_block.IN  :=IN;
	func_block.PT  :=PT;
	func_block();
	Q := func_block.Q;

END_PROGRAM

CONFIGURATION Config0
	RESOURCE Res0 ON PLC
		TASK task0(INTERVAL := T#20ms,PRIORITY := 0);
		PROGRAM instance0 WITH task0 : program0;
	END_RESOURCE
END_CONFIGURATION

(* ---- TN_FRAMEWORK.ST ---- *)
TYPE
  bya_TN_CHAR:       	ARRAY [0..1919] OF BYTE;
  bya_TN_BACKUP:     	ARRAY [0..1919] OF BYTE;
  bya_TN_COLOR:      	ARRAY [0..1919] OF BYTE;
  bya_TN_Line_Update:	ARRAY [0..23]   OF BOOL;

  us_TN_SCREEN :
  STRUCT
		bya_CHAR:			bya_TN_CHAR;
		bya_COLOR:			bya_TN_COLOR;
		bya_BACKUP:			bya_TN_BACKUP;
		bya_Line_Update:	bya_TN_Line_Update;

		by_Input_Exten_Code:    BYTE;
		by_Input_ASCII_Code:    BYTE;
		bo_Input_ASCII_IsNum:   BOOL;
		in_Page_Number:        	INT;
		in_Cursor_X:           	INT;
		in_Cursor_Y:           	INT;
		in_EOS_Offset:         	INT;
		by_Clear_Screen_Attr:  	BYTE;
		bo_Clear_Screen:       	BOOL;
		bo_Modal_Dialog:       	BOOL;
		bo_Menue_Bar_Dialog:   	BOOL;

  END_STRUCT;
END_TYPE

TYPE
  oscat_NW_BUF_LONG  : ARRAY [0..4095] OF BYTE;

  oscat_NETWORK_BUFFER :
  STRUCT
    SIZE   : UINT;
    BUFFER : oscat_NW_BUF_LONG;
  END_STRUCT;
END_TYPE

FUNCTION ISC_NUM:BOOL

	VAR_INPUT
		IN :	BYTE;
	END_VAR

	ISC_NUM := IN > BYTE#47 AND IN < BYTE#58;

END_FUNCTION

FUNCTION_BLOCK TN_RECEIVE_Block

  VAR_IN_OUT
    R_BUF :	oscat_NETWORK_BUFFER;
    Xus_TN_SCREEN :	us_TN_SCREEN;
  END_VAR

  VAR
    REQ_Size :	UINT;
    REQ1 :	BYTE;
    REQ2 :	BYTE;
    REQ3 :	BYTE;
  END_VAR

  Xus_TN_SCREEN.by_Input_ASCII_Code := BYTE#00;
  Xus_TN_SCREEN.by_Input_Exten_Code := BYTE#00;

  IF R_BUF.SIZE > UINT#0 THEN
    REQ_Size := R_BUF.SIZE;
    REQ1 := R_BUF.BUFFER[0];
    REQ2 := R_BUF.BUFFER[1];
    REQ3 := R_BUF.BUFFER[2];

    IF REQ1 = BYTE#27 AND REQ_Size >= UINT#3 THEN
      IF REQ2 = BYTE#91 THEN
        IF (REQ3 >= BYTE#65 AND REQ3 <= BYTE#68) OR (REQ3 = BYTE#72) OR (REQ3 = BYTE#75) THEN
          Xus_TN_SCREEN.by_Input_Exten_Code := REQ3;
        END_IF;
      ELSIF REQ2 = BYTE#79 THEN
        IF REQ3 >= BYTE#80 AND REQ3 <= BYTE#83 THEN
          Xus_TN_SCREEN.by_Input_Exten_Code := REQ3;
        END_IF;
      END_IF;
    ELSIF REQ1 >= BYTE#32 AND REQ1 <= BYTE#126 THEN
    Xus_TN_SCREEN.by_Input_ASCII_Code := REQ1;
      Xus_TN_SCREEN.bo_Input_ASCII_IsNum := ISC_NUM(REQ1);
    ELSIF REQ1 = BYTE#8 OR REQ1 = BYTE#9 OR REQ1 = BYTE#13 OR REQ1 = BYTE#27 THEN
    Xus_TN_SCREEN.by_Input_Exten_Code := REQ1;
    END_IF;

    R_BUF.SIZE := UINT#00;
  END_IF;

END_FUNCTION_BLOCK

TYPE
  oscat_IP_FIFO128_DATA  : ARRAY [1..128] OF BYTE;
  oscat_Mailbox  : ARRAY [1..16] OF BYTE;

  oscat_IP_FIFO_DATA :
  STRUCT
    X       : oscat_IP_FIFO128_DATA; (* IP_ID FIFO Speicher          *)
    Y       : oscat_IP_FIFO128_DATA; (* IP_ID Z�hler                 *)
    ID      : BYTE;                  (* h�chste vergabene id         *)
    MAX_ID  : BYTE;                  (* maximal Anmeldungen pro ID   *)
    INIT    : BOOL;                  (* Initialisierung durchgef�hrt *)
    EMPTY   : BOOL;                  (* FIFO leer                    *)
    FULL    : BOOL;                  (* FIFO voll                    *)
    TOP     : INT;                   (* maximale anzahl in FIFO      *)
    NW      : INT;                   (* Schreibzeiger                *)
    NR      : INT;                   (* Lesezeiger                   *)
  END_STRUCT;

  oscat_IP_C:
  STRUCT
    C_MODE:			BYTE;          		(*W Mode: TCP/UCP AKTIV/PASSIV                               *)
    C_PORT:         WORD;          		(*W Portnummer                                               *)
    C_IP:           DWORD;         		(*W IP-Adresse gepackt wwxxyyzz = www.xxx.yyy.zzz            *)
    C_STATE:        BYTE;          		(*R Verbindungsstatus ON/OFF + Flanke ON/OFF                 *)
    C_ENABLE:       BOOL;          		(*W Freigabe f�r Connect                                     *)
    R_OBSERVE:      BOOL;          		(*W Empfang ueberwachen                                      *)
    TIME_RESET:     BOOL;          		(*W Alle Timer ruecksetzen                                   *)
    ERROR:          DWORD;         		(*R vvwwxxyy (vv = CON_ERROR, ww = SEN_ERROR, xx = REC_ERROR *)
    FIFO:           oscat_IP_FIFO_DATA; (*I IP FIFO Struktur                                         *)
    MAILBOX:		oscat_Mailbox;		(*I Mailbox: Datenbereich f�r Bausteindatenaustausch         *)
    END_STRUCT;
END_TYPE

FUNCTION INT_TO_BCDC:BYTE

	VAR_INPUT
		IN :	INT;
	END_VAR

	INT_TO_BCDC := SHL(INT_TO_BYTE(IN / INT#10),4) OR INT_TO_BYTE(in MOD INT#10);

END_FUNCTION

FUNCTION_BLOCK TN_SEND_ROWS_Block

  VAR_IN_OUT
    IP_C :	oscat_IP_C;
    S_BUF :	oscat_NETWORK_BUFFER;
    Xus_TN_SCREEN :	us_TN_SCREEN;
  END_VAR

  VAR_INPUT
    S_BUF_SIZE :	INT;
  END_VAR

  VAR
    in_Line_Count :	INT;
    in_Col_Count :	INT;
    in_Last_Row_Index :	INT;
    bo_Break_Loop :	BOOL;
    in_Row_Count :	INT;
    in_Offset :	INT;
    in_Write_Index :	INT;
    in_Write_Index_Backup :	INT;
    by_Cur_Color :	BYTE;
    by_last_Color :	BYTE;
    in_Write_Stop :	INT;
  END_VAR

  IF (IP_C.C_STATE < BYTE#127 OR S_BUF.SIZE > UINT#0) THEN
    RETURN;
  END_IF;

  in_Write_Index := UINT_TO_INT(S_BUF.SIZE) - 1;

  in_Write_Index_Backup := in_Write_Index;

  IF (IP_C.C_STATE = BYTE#254) OR (Xus_TN_SCREEN.bo_Clear_Screen) THEN

    Xus_TN_SCREEN.bo_Clear_Screen := FALSE;

    FOR in_Line_Count := INT#00 TO INT#23 DO
      Xus_TN_SCREEN.bya_Line_Update[in_Line_Count] := TRUE;
    END_FOR;

    in_Write_Index := in_Write_Index + INT#1;
    S_BUF.BUFFER[in_Write_Index] := BYTE#16#1B;
    in_Write_Index := in_Write_Index + INT#1;
    S_BUF.BUFFER[in_Write_Index] := BYTE#16#5B;
    in_Write_Index := in_Write_Index + INT#1;
    S_BUF.BUFFER[in_Write_Index] := BYTE#16#30;
    in_Write_Index := in_Write_Index + INT#1;
    S_BUF.BUFFER[in_Write_Index] := BYTE#16#3B;
    in_Write_Index := in_Write_Index + INT#1;
    S_BUF.BUFFER[in_Write_Index] := BYTE#16#33;

    in_Write_Index := in_Write_Index + INT#1;
    S_BUF.BUFFER[in_Write_Index] := (SHR(Xus_TN_SCREEN.by_Clear_Screen_Attr,4) OR BYTE#16#30);

    in_Write_Index := in_Write_Index + INT#1;
    S_BUF.BUFFER[in_Write_Index] := BYTE#16#3B;
    in_Write_Index := in_Write_Index + INT#1;
    S_BUF.BUFFER[in_Write_Index] := BYTE#16#34;

    in_Write_Index := in_Write_Index + INT#1;
    S_BUF.BUFFER[in_Write_Index] := ((Xus_TN_SCREEN.by_Clear_Screen_Attr AND BYTE#16#07) OR BYTE#16#30);

    in_Write_Index := in_Write_Index + INT#1;
    S_BUF.BUFFER[in_Write_Index] := BYTE#16#6D;

    in_Write_Index := in_Write_Index + INT#1;
    S_BUF.BUFFER[in_Write_Index] := BYTE#16#1B;
    in_Write_Index := in_Write_Index + INT#1;
    S_BUF.BUFFER[in_Write_Index] := BYTE#16#5B;
    in_Write_Index := in_Write_Index + INT#1;
    S_BUF.BUFFER[in_Write_Index] := BYTE#16#32;
    in_Write_Index := in_Write_Index + INT#1;
    S_BUF.BUFFER[in_Write_Index] := BYTE#16#4A;

    in_Write_Index := in_Write_Index + INT#1;
    S_BUF.BUFFER[in_Write_Index] := BYTE#16#1B;
    in_Write_Index := in_Write_Index + INT#1;
    S_BUF.BUFFER[in_Write_Index] := BYTE#16#5B;
    in_Write_Index := in_Write_Index + INT#1;
    S_BUF.BUFFER[in_Write_Index] := BYTE#16#3F;
    in_Write_Index := in_Write_Index + INT#1;
    S_BUF.BUFFER[in_Write_Index] := BYTE#16#37;
    in_Write_Index := in_Write_Index + INT#1;
    S_BUF.BUFFER[in_Write_Index] := BYTE#16#6C;

  END_IF;

  in_Last_Row_Index := INT#0;
  bo_Break_Loop := FALSE;
  in_Write_Stop := S_BUF_SIZE-20;

  FOR in_Line_Count := 0 TO 23 DO

    in_Offset := in_Row_Count * INT#80;

    IF (Xus_TN_SCREEN.bya_Line_Update[in_Row_Count] = TRUE) THEN

      in_Write_Index := in_Write_Index + INT#1;
      S_BUF.BUFFER[in_Write_Index] := BYTE#16#1B;
      in_Write_Index := in_Write_Index + INT#1;
      S_BUF.BUFFER[in_Write_Index] := BYTE#16#5B;

      in_Write_Index := in_Write_Index + INT#1;
      S_BUF.BUFFER[in_Write_Index] :=
        SHR(INT_TO_BCDC(in_Row_Count + INT#1),INT#4) OR BYTE#16#30;

      in_Write_Index := in_Write_Index + INT#1;
      S_BUF.BUFFER[in_Write_Index] :=
        (INT_TO_BCDC(in_Row_Count + INT#1) AND BYTE#16#0F) OR BYTE#16#30;

      in_Write_Index := in_Write_Index + INT#1;
      S_BUF.BUFFER[in_Write_Index] := BYTE#16#3B;
      in_Write_Index := in_Write_Index + INT#1;
      S_BUF.BUFFER[in_Write_Index] := BYTE#16#31;
      in_Write_Index := in_Write_Index + INT#1;
      S_BUF.BUFFER[in_Write_Index] := BYTE#16#48;

      FOR in_Col_Count := 0 TO 79 DO

        by_Cur_Color := Xus_TN_SCREEN.bya_COLOR[in_Offset];
        IF (by_Cur_Color <> by_last_Color) OR (in_Col_Count = INT#00) THEN

          in_Write_Index := in_Write_Index + INT#1;
          S_BUF.BUFFER[in_Write_Index] := BYTE#16#1B;

          in_Write_Index := in_Write_Index + INT#1;
          S_BUF.BUFFER[in_Write_Index] := BYTE#16#5B;

          IF  (((by_Cur_Color AND BYTE#2#10001000) XOR (by_last_Color AND BYTE#2#10001000)) <> BYTE#00) OR (in_Col_Count = 0) THEN

            in_Write_Index := in_Write_Index + INT#1;
            S_BUF.BUFFER[in_Write_Index] := BYTE#16#30;
            in_Write_Index := in_Write_Index + INT#1;
            S_BUF.BUFFER[in_Write_Index] := BYTE#16#3B;

            IF (by_Cur_Color AND BYTE#2#00001000) = BYTE#2#00000000 THEN

              in_Write_Index := in_Write_Index + INT#1;
              S_BUF.BUFFER[in_Write_Index] := BYTE#16#31;
              in_Write_Index := in_Write_Index + INT#1;
              S_BUF.BUFFER[in_Write_Index] := BYTE#16#3B;

            END_IF;

            IF (by_Cur_Color AND BYTE#2#10000000) = BYTE#2#10000000 THEN

              in_Write_Index := in_Write_Index + INT#1;
              S_BUF.BUFFER[in_Write_Index] := BYTE#16#35;
              in_Write_Index := in_Write_Index + INT#1;
              S_BUF.BUFFER[in_Write_Index] := BYTE#16#3B;

            END_IF;

          END_IF;

          in_Write_Index := in_Write_Index + INT#1;
          S_BUF.BUFFER[in_Write_Index] := BYTE#16#33;

          in_Write_Index := in_Write_Index + INT#1;
          S_BUF.BUFFER[in_Write_Index] := ((SHR(by_Cur_Color,4) AND BYTE#2#00000111) OR BYTE#16#30);

          in_Write_Index := in_Write_Index + INT#1;
          S_BUF.BUFFER[in_Write_Index] := BYTE#16#3B;

          in_Write_Index := in_Write_Index + INT#1;
          S_BUF.BUFFER[in_Write_Index] := BYTE#16#34;

          in_Write_Index := in_Write_Index + INT#1;
          S_BUF.BUFFER[in_Write_Index] := ((by_Cur_Color AND BYTE#2#00000111) OR BYTE#16#30);

          in_Write_Index := in_Write_Index + INT#1;
          S_BUF.BUFFER[in_Write_Index] := BYTE#16#6D;

          by_last_Color := by_Cur_Color;

        END_IF;

        IF (in_Write_Index > in_Write_Stop) THEN

          bo_Break_Loop := TRUE;
          EXIT;

        END_IF;

        in_Write_Index := in_Write_Index + INT#1;
        S_BUF.BUFFER[in_Write_Index] := Xus_TN_SCREEN.bya_CHAR[in_Offset];

        in_Offset := in_Offset + INT#01;
      END_FOR;

      IF (bo_Break_Loop = TRUE) THEN

        in_Write_Index := in_Last_Row_Index;

        EXIT;
      END_IF;

      in_Last_Row_Index := in_Write_Index;
      Xus_TN_SCREEN.bya_Line_Update[in_Row_Count] := FALSE;

    END_IF;

    in_Row_Count := in_Row_Count + INT#01;

    IF (in_Row_Count > INT#23) THEN
      in_Row_Count := INT#00;
    END_IF;

  END_FOR;

  IF (bo_Break_Loop = FALSE) THEN

    in_Row_Count := INT#00;

  END_IF;

  IF (in_Write_Index <> in_Write_Index_Backup) THEN

    in_Write_Index := in_Write_Index + INT#1;
    S_BUF.BUFFER[in_Write_Index] := BYTE#16#1B;
    in_Write_Index := in_Write_Index + INT#1;
    S_BUF.BUFFER[in_Write_Index] := BYTE#16#5B;

    in_Write_Index := in_Write_Index + INT#1;
    S_BUF.BUFFER[in_Write_Index] := SHR(INT_TO_BCDC(Xus_TN_SCREEN.in_Cursor_Y + 1),INT#4) OR BYTE#16#30;

    in_Write_Index := in_Write_Index + INT#1;
    S_BUF.BUFFER[in_Write_Index] := (INT_TO_BCDC(Xus_TN_SCREEN.in_Cursor_Y + 1) AND BYTE#16#0F) OR BYTE#16#30;

    in_Write_Index := in_Write_Index + INT#1;
    S_BUF.BUFFER[in_Write_Index] := BYTE#16#3B;

    in_Write_Index := in_Write_Index + INT#1;
    S_BUF.BUFFER[in_Write_Index] := SHR(INT_TO_BCDC(Xus_TN_SCREEN.in_Cursor_X + 1),INT#4) OR BYTE#16#30;

    in_Write_Index := in_Write_Index + INT#1;
    S_BUF.BUFFER[in_Write_Index] := (INT_TO_BCDC(Xus_TN_SCREEN.in_Cursor_X + 1) AND BYTE#16#0F) OR BYTE#16#30;

    in_Write_Index := in_Write_Index + INT#1;
    S_BUF.BUFFER[in_Write_Index] := BYTE#16#48;

  END_IF;

  S_BUF.SIZE := INT_TO_UINT(in_Write_Index + 1);

END_FUNCTION_BLOCK

FUNCTION_BLOCK TN_FRAMEWORK_Block

	VAR_IN_OUT
		us_TN_INPUT_CONTROL :	us_TN_INPUT_CONTROL;
		us_TN_SCREEN :	us_TN_SCREEN;
		us_TN_MENU :	us_TN_MENU;
		S_BUF :	oscat_NETWORK_BUFFER;
		R_BUF :	oscat_NETWORK_BUFFER;
		IP_C :	oscat_IP_C;
	END_VAR

	VAR
		FB_IP_CONTROL :	IP_CONTROL;
		FB_TN_INPUT_CONTROL :	TN_INPUT_CONTROL;
		FB_TN_INPUT_MENU_BAR :	TN_INPUT_MENU_BAR;
		FB_TN_RECEIVE :	TN_RECEIVE_Block;
		FB_TN_SEND_ROWS :	TN_SEND_ROWS_Block;
		t :	TON;
	END_VAR

	IF (NOT IP_C.C_ENABLE) THEN

	IP_C.C_PORT     := WORD#23;
	IP_C.C_IP       := DWORD#00;
	IP_C.C_MODE     := BYTE#4;
	IP_C.TIME_RESET := TRUE;
	IP_C.C_ENABLE   := TRUE;
	IP_C.R_OBSERVE  := FALSE;

	END_IF;

	t(IN:= IP_C.ERROR > DWORD#0, PT:=T#5s);
	IF t.Q THEN
		IP_C.TIME_RESET := TRUE;
	END_IF;

	FB_TN_INPUT_MENU_BAR.Xus_TN_MENU    := us_TN_MENU;
	FB_TN_INPUT_MENU_BAR.Xus_TN_SCREEN  := us_TN_SCREEN;
	FB_TN_INPUT_MENU_BAR();
	us_TN_MENU   := FB_TN_INPUT_MENU_BAR.Xus_TN_MENU;
	us_TN_SCREEN := FB_TN_INPUT_MENU_BAR.Xus_TN_SCREEN;

	FB_TN_INPUT_CONTROL.Xus_TN_SCREEN        := us_TN_SCREEN;
	FB_TN_INPUT_CONTROL.Xus_TN_INPUT_CONTROL := us_TN_INPUT_CONTROL;
	FB_TN_INPUT_CONTROL();
	us_TN_SCREEN        := FB_TN_INPUT_CONTROL.Xus_TN_SCREEN;
	us_TN_INPUT_CONTROL := FB_TN_INPUT_CONTROL.Xus_TN_INPUT_CONTROL;

	FB_TN_SEND_ROWS.IP_C          := IP_C;
	FB_TN_SEND_ROWS.S_BUF         := S_BUF;
	FB_TN_SEND_ROWS.Xus_TN_SCREEN := us_TN_SCREEN;
	FB_TN_SEND_ROWS.S_BUF_SIZE    := 4096;
	FB_TN_SEND_ROWS();
	IP_C         := FB_TN_SEND_ROWS.IP_C;
	S_BUF        := FB_TN_SEND_ROWS.S_BUF;
	us_TN_SCREEN := FB_TN_SEND_ROWS.Xus_TN_SCREEN;

	FB_IP_CONTROL.IP_C     := IP_C;
	FB_IP_CONTROL.S_BUF    := S_BUF;
	FB_IP_CONTROL.R_BUF    := R_BUF;
	FB_IP_CONTROL.IP       := DWORD#00;
	FB_IP_CONTROL.PORT     := WORD#00;
	FB_IP_CONTROL.TIME_OUT := T#2s;
	FB_IP_CONTROL();
	IP_C  := FB_IP_CONTROL.IP_C;
	S_BUF := FB_IP_CONTROL.S_BUF;
	R_BUF := FB_IP_CONTROL.R_BUF;

	FB_TN_RECEIVE.R_BUF := R_BUF;
	FB_TN_RECEIVE.Xus_TN_SCREEN := us_TN_SCREEN;
	FB_TN_RECEIVE();
	R_BUF := FB_TN_RECEIVE.R_BUF;
	us_TN_SCREEN := FB_TN_RECEIVE.Xus_TN_SCREEN;

END_FUNCTION_BLOCK

PROGRAM program0
	VAR
		R_BUF :	oscat_NETWORK_BUFFER;
    Xus_TN_SCREEN :	us_TN_SCREEN;

		func_block : TN_RECEIVE_Block;
	END_VAR
	func_block.R_BUF := R_BUF;
	func_block.Xus_TN_SCREEN := Xus_TN_SCREEN;

	func_block();
  R_BUF  := func_block.R_BUF;
	Xus_TN_SCREEN  := func_block.Xus_TN_SCREEN;
END_PROGRAM

CONFIGURATION Config0
	RESOURCE Res0 ON PLC
		TASK task0(INTERVAL := T#20ms,PRIORITY := 0);
		PROGRAM instance0 WITH task0 : program0;
	END_RESOURCE
END_CONFIGURATION

(* ---- TN_INPUT_CONTROL.ST ---- *)
FUNCTION_BLOCK TN_INPUT_CONTROL

  VAR_IN_OUT
    Xus_TN_SCREEN :	us_TN_SCREEN;
    Xus_TN_INPUT_CONTROL :	us_TN_INPUT_CONTROL;
  END_VAR

  VAR
    FB_TN_INPUT_SELECT_POPUP :	TN_INPUT_SELECT_POPUP;
  END_VAR

  VAR
    FB_TN_INPUT_SELECT_TEXT :	TN_INPUT_SELECT_TEXT;
    FB_TN_SC_WRITE_C :	TN_SC_WRITE_C;
    FB_TN_INPUT_EDIT_LINE :	TN_INPUT_EDIT_LINE;
  END_VAR

  VAR
    in_index :	INT;
    in_Scroll_Offset :	INT;
    in_Focus_new :	INT;
    in_Focus_alt :	INT;
    bo_Tool_Tip_Update :	BOOL;
  END_VAR

  IF (Xus_TN_INPUT_CONTROL.bo_Enable = FALSE) OR (Xus_TN_SCREEN.bo_Menue_Bar_Dialog = TRUE) THEN
    RETURN;
  END_IF;

  IF (Xus_TN_INPUT_CONTROL.bo_Reset_Fokus = TRUE) THEN

    Xus_TN_INPUT_CONTROL.bo_Reset_Fokus := FALSE;

    FOR in_index := INT#01 TO Xus_TN_INPUT_CONTROL.in_Count DO
      Xus_TN_INPUT_CONTROL.usa_TN_INPUT_CONTROL_DATA[in_index].bo_Focus := FALSE;
    END_FOR;

    IF (Xus_TN_INPUT_CONTROL.in_Count >= INT#01) THEN

      Xus_TN_INPUT_CONTROL.usa_TN_INPUT_CONTROL_DATA[1].bo_Focus := TRUE;
      Xus_TN_INPUT_CONTROL.in_Focus_at := INT#01;

    END_IF;

    Xus_TN_INPUT_CONTROL.bo_Update_all := TRUE;

  END_IF;

  IF (Xus_TN_SCREEN.bo_Modal_Dialog = FALSE) THEN

    IF (Xus_TN_SCREEN.by_Input_Exten_Code = BYTE#09) THEN

      in_Scroll_Offset := INT#01;

    ELSIF (Xus_TN_SCREEN.by_Input_Exten_Code = BYTE#65) THEN

      in_Scroll_Offset := INT#-01;

    ELSIF (Xus_TN_SCREEN.by_Input_Exten_Code = BYTE#66) THEN

      in_Scroll_Offset := INT#01;

    END_IF;
  END_IF;

  IF (in_Scroll_Offset <> INT#00) THEN

    Xus_TN_INPUT_CONTROL.in_Focus_at:=LIMIT_INT(INT#01,Xus_TN_INPUT_CONTROL.in_Focus_at,Xus_TN_INPUT_CONTROL.in_Count);

    in_Focus_new := Xus_TN_INPUT_CONTROL.in_Focus_at + in_Scroll_Offset;

    IF (in_Focus_new > Xus_TN_INPUT_CONTROL.in_Count) THEN
      in_Focus_new := INT#1;
    END_IF;

    IF (in_Focus_new < INT#01) THEN
      in_Focus_new := Xus_TN_INPUT_CONTROL.in_Count;
    END_IF;

    in_Focus_alt := Xus_TN_INPUT_CONTROL.in_Focus_at;

    Xus_TN_INPUT_CONTROL.usa_TN_INPUT_CONTROL_DATA[in_Focus_alt].bo_Focus := FALSE;
    Xus_TN_INPUT_CONTROL.usa_TN_INPUT_CONTROL_DATA[in_Focus_alt].bo_Update_Input := TRUE;

    Xus_TN_INPUT_CONTROL.usa_TN_INPUT_CONTROL_DATA[in_Focus_new].bo_Focus  := TRUE;
    Xus_TN_INPUT_CONTROL.usa_TN_INPUT_CONTROL_DATA[in_Focus_new].bo_Update_Input := TRUE;

    Xus_TN_INPUT_CONTROL.in_Focus_at := in_Focus_new;

    bo_Tool_Tip_Update := TRUE;
    in_Scroll_Offset := INT#00;

  END_IF;

  IF (Xus_TN_INPUT_CONTROL.bo_Update_all = TRUE) THEN
    FOR in_index := 1 TO Xus_TN_INPUT_CONTROL.in_Count DO
      Xus_TN_INPUT_CONTROL.usa_TN_INPUT_CONTROL_DATA[in_index].bo_Update_All := TRUE;
    END_FOR;
    Xus_TN_INPUT_CONTROL.bo_Update_all := FALSE;
    bo_Tool_Tip_Update := TRUE;
  END_IF;

  FOR in_index := 1 TO Xus_TN_INPUT_CONTROL.in_Count DO

    IF (Xus_TN_INPUT_CONTROL.usa_TN_INPUT_CONTROL_DATA[in_index].in_Type > INT#00) THEN

      IF (Xus_TN_INPUT_CONTROL.usa_TN_INPUT_CONTROL_DATA[in_index].bo_Focus = TRUE) THEN

        Xus_TN_INPUT_CONTROL.usa_TN_INPUT_CONTROL_DATA[in_index].by_Input_ASCII_Code  := Xus_TN_SCREEN.by_Input_ASCII_Code;
        Xus_TN_INPUT_CONTROL.usa_TN_INPUT_CONTROL_DATA[in_index].by_Input_Exten_Code  := Xus_TN_SCREEN.by_Input_Exten_Code;
        Xus_TN_INPUT_CONTROL.usa_TN_INPUT_CONTROL_DATA[in_index].bo_Input_ASCII_IsNum := Xus_TN_SCREEN.bo_Input_ASCII_IsNum;

        IF (bo_Tool_Tip_Update = TRUE) THEN

          FB_TN_SC_WRITE_C.Iin_Y          := Xus_TN_INPUT_CONTROL.in_ToolTip_Y;
          FB_TN_SC_WRITE_C.Iin_X          := Xus_TN_INPUT_CONTROL.in_ToolTip_X;
          FB_TN_SC_WRITE_C.Iby_ATTR       := Xus_TN_INPUT_CONTROL.by_ToolTip_Attr;
          FB_TN_SC_WRITE_C.Iin_OPTION     := INT#02;
          FB_TN_SC_WRITE_C.Iin_LENGTH     := Xus_TN_INPUT_CONTROL.in_ToolTip_Size;
          FB_TN_SC_WRITE_C.Ist_STRING     := Xus_TN_INPUT_CONTROL.usa_TN_INPUT_CONTROL_DATA[in_index].st_Input_ToolTip;
          FB_TN_SC_WRITE_C.Xus_TN_SCREEN  := Xus_TN_SCREEN;
          FB_TN_SC_WRITE_C();
          Xus_TN_SCREEN := FB_TN_SC_WRITE_C.Xus_TN_SCREEN;

          bo_Tool_Tip_Update := FALSE;

        END_IF;

      END_IF;

      CASE Xus_TN_INPUT_CONTROL.usa_TN_INPUT_CONTROL_DATA[in_index].in_Type OF

      1:
        FB_TN_INPUT_EDIT_LINE.Xus_TN_INPUT_CONTROL_DATA := Xus_TN_INPUT_CONTROL.usa_TN_INPUT_CONTROL_DATA[in_index];
        FB_TN_INPUT_EDIT_LINE.Xus_TN_SCREEN             := Xus_TN_SCREEN;
        FB_TN_INPUT_EDIT_LINE();
        Xus_TN_INPUT_CONTROL.usa_TN_INPUT_CONTROL_DATA[in_index]  := FB_TN_INPUT_EDIT_LINE.Xus_TN_INPUT_CONTROL_DATA;
        Xus_TN_SCREEN                                             := FB_TN_INPUT_EDIT_LINE.Xus_TN_SCREEN;

      2:
        FB_TN_INPUT_SELECT_TEXT.Xus_TN_INPUT_CONTROL_DATA := Xus_TN_INPUT_CONTROL.usa_TN_INPUT_CONTROL_DATA[in_index];
        FB_TN_INPUT_SELECT_TEXT.Xus_TN_SCREEN             := Xus_TN_SCREEN;
        FB_TN_INPUT_SELECT_TEXT();
        Xus_TN_INPUT_CONTROL.usa_TN_INPUT_CONTROL_DATA[in_index] := FB_TN_INPUT_SELECT_TEXT.Xus_TN_INPUT_CONTROL_DATA;
        Xus_TN_SCREEN                                            := FB_TN_INPUT_SELECT_TEXT.Xus_TN_SCREEN;
      3:
        FB_TN_INPUT_SELECT_POPUP.Xus_TN_INPUT_CONTROL_DATA := Xus_TN_INPUT_CONTROL.usa_TN_INPUT_CONTROL_DATA[in_index];
        FB_TN_INPUT_SELECT_POPUP.Xus_TN_SCREEN             := Xus_TN_SCREEN;
        FB_TN_INPUT_SELECT_POPUP();
        Xus_TN_INPUT_CONTROL.usa_TN_INPUT_CONTROL_DATA[in_index] := FB_TN_INPUT_SELECT_POPUP.Xus_TN_INPUT_CONTROL_DATA;
        Xus_TN_SCREEN                                            := FB_TN_INPUT_SELECT_POPUP.Xus_TN_SCREEN;

      END_CASE;

      IF (Xus_TN_INPUT_CONTROL.usa_TN_INPUT_CONTROL_DATA[in_index].bo_Focus = TRUE) THEN

        Xus_TN_SCREEN.in_Cursor_X := Xus_TN_INPUT_CONTROL.usa_TN_INPUT_CONTROL_DATA[in_index].in_Cursor_X;
        Xus_TN_SCREEN.in_Cursor_Y := Xus_TN_INPUT_CONTROL.usa_TN_INPUT_CONTROL_DATA[in_index].in_Cursor_Y;

      END_IF;
    END_IF;
  END_FOR;

END_FUNCTION_BLOCK

(* ---- TN_INPUT_EDIT_LINE.ST ---- *)
FUNCTION_BLOCK TN_INPUT_EDIT_LINE

  VAR
    in_count :	INT;
    in_Count_End :	INT;
    in_CursorOffset :	INT;
    by_Attr :	BYTE;
    st_String :	STRING;
    bo_Pos_Found :	BOOL;
    st_CHAR :	oscat_STRING1;
    in_old_charpos :	INT;
  END_VAR

  VAR
    FB_TN_SC_WRITE :	TN_SC_WRITE;
    CHR_TO_STRING :	CHR_TO_STRING;
    FB_TRIME :	TRIME;
  END_VAR

  VAR_IN_OUT
    Xus_TN_SCREEN :	us_TN_SCREEN;
    Xus_TN_INPUT_CONTROL_DATA :	us_TN_INPUT_CONTROL_DATA;
  END_VAR

  in_CursorOffset := INT#0;

  IF Xus_TN_INPUT_CONTROL_DATA.bo_Focus = TRUE THEN

    IF Xus_TN_INPUT_CONTROL_DATA.by_Input_ASCII_Code > BYTE#0 THEN

      IF (Xus_TN_INPUT_CONTROL_DATA.bo_Input_Only_Num = TRUE AND Xus_TN_INPUT_CONTROL_DATA.bo_Input_ASCII_IsNum = TRUE)
        OR (Xus_TN_INPUT_CONTROL_DATA.bo_Input_Only_Num = FALSE) THEN

        CHR_TO_STRING(C:=Xus_TN_INPUT_CONTROL_DATA.by_Input_ASCII_Code);
        st_CHAR:=CHR_TO_STRING.CHR_TO_STRING;

        Xus_TN_INPUT_CONTROL_DATA.st_Input_Data := REPLACE(Xus_TN_INPUT_CONTROL_DATA.st_Input_Data,
        st_CHAR,INT#1,Xus_TN_INPUT_CONTROL_DATA.in_Cursor_Pos);

        in_CursorOffset := INT#1;
        Xus_TN_INPUT_CONTROL_DATA.bo_Update_Input := TRUE;
      END_IF;

    END_IF;

    CASE _BYTE_TO_INT(Xus_TN_INPUT_CONTROL_DATA.by_Input_Exten_Code) OF

    67:
      in_CursorOffset := INT#1;

    68:
      in_CursorOffset := INT#-1;

    08:
      Xus_TN_INPUT_CONTROL_DATA.st_Input_Data :=REPLACE(Xus_TN_INPUT_CONTROL_DATA.st_Input_Data,' ',INT#1,Xus_TN_INPUT_CONTROL_DATA.in_Cursor_Pos);
      Xus_TN_INPUT_CONTROL_DATA.bo_Update_Input := TRUE;
      in_CursorOffset := INT#-1;

    13:
      IF LEN(Xus_TN_INPUT_CONTROL_DATA.st_Input_Mask) > INT#00 THEN
        Xus_TN_INPUT_CONTROL_DATA.st_Input_String := Xus_TN_INPUT_CONTROL_DATA.st_Input_Data;

        FB_TRIME(str:=Xus_TN_INPUT_CONTROL_DATA.st_Input_String);
        Xus_TN_INPUT_CONTROL_DATA.st_Input_String:=FB_TRIME.TRIME;

        Xus_TN_INPUT_CONTROL_DATA.bo_Input_Entered := TRUE;

        Xus_TN_INPUT_CONTROL_DATA.st_Input_Data := Xus_TN_INPUT_CONTROL_DATA.st_Input_Mask;

        Xus_TN_INPUT_CONTROL_DATA.in_Cursor_Pos := INT#1;
        Xus_TN_INPUT_CONTROL_DATA.bo_Update_Input := TRUE;

        st_CHAR := MID(Xus_TN_INPUT_CONTROL_DATA.st_Input_Mask,1,Xus_TN_INPUT_CONTROL_DATA.in_Cursor_Pos);
        IF NE_STRING(st_CHAR,' ') THEN
          in_CursorOffset := INT#1;
        END_IF;
      END_IF;
    END_CASE;
  END_IF;

  IF (in_CursorOffset > INT#0) OR (Xus_TN_INPUT_CONTROL_DATA.in_Cursor_Pos = INT#0) THEN
    bo_Pos_Found := FALSE;

    in_Count     := Xus_TN_INPUT_CONTROL_DATA.in_Cursor_Pos + INT#1;
    in_Count_End := LEN(Xus_TN_INPUT_CONTROL_DATA.st_Input_Mask);

    WHILE (in_count <= in_Count_End) AND (bo_Pos_Found = FALSE)  DO

      st_CHAR := MID(Xus_TN_INPUT_CONTROL_DATA.st_Input_Mask,1,in_count);
      IF EQ_STRING(st_CHAR,' ') THEN
        Xus_TN_INPUT_CONTROL_DATA.in_Cursor_Pos := in_count;
        Xus_TN_INPUT_CONTROL_DATA.bo_Update_Input := TRUE;
        bo_Pos_Found := TRUE;
      END_IF;

      in_count := in_count + INT#1;

    END_WHILE;

  END_IF;

  IF in_CursorOffset < INT#0 THEN
    bo_Pos_Found := FALSE;

    in_Count     := Xus_TN_INPUT_CONTROL_DATA.in_Cursor_Pos - INT#01;
    in_Count_End := INT#1;

    WHILE (in_count >= in_Count_End) AND (bo_Pos_Found = FALSE) DO

      st_CHAR := MID(Xus_TN_INPUT_CONTROL_DATA.st_Input_Mask,1,in_count);
      IF EQ_STRING(st_CHAR,' ') THEN
        Xus_TN_INPUT_CONTROL_DATA.in_Cursor_Pos := in_count;
        Xus_TN_INPUT_CONTROL_DATA.bo_Update_Input := TRUE;
        bo_Pos_Found := TRUE;
      END_IF;

      in_count := in_count - INT#1;
    END_WHILE;

  END_IF;

  IF Xus_TN_INPUT_CONTROL_DATA.in_Cursor_Pos > LEN(Xus_TN_INPUT_CONTROL_DATA.st_Input_Data) THEN
    Xus_TN_INPUT_CONTROL_DATA.in_Cursor_Pos := LEN(Xus_TN_INPUT_CONTROL_DATA.st_Input_Data);
    Xus_TN_INPUT_CONTROL_DATA.bo_Update_Input := TRUE;
  END_IF;

  IF Xus_TN_INPUT_CONTROL_DATA.in_Cursor_Pos < INT#1 THEN
    Xus_TN_INPUT_CONTROL_DATA.in_Cursor_Pos := INT#1;
    Xus_TN_INPUT_CONTROL_DATA.bo_Update_Input := TRUE;
  END_IF;
  IF (Xus_TN_INPUT_CONTROL_DATA.bo_Update_Input = TRUE) OR (Xus_TN_INPUT_CONTROL_DATA.bo_Update_All = TRUE) THEN

    IF (Xus_TN_INPUT_CONTROL_DATA.bo_Update_All = TRUE) THEN

      IF (Xus_TN_INPUT_CONTROL_DATA.in_Title_X_Offset = INT#00) AND (Xus_TN_INPUT_CONTROL_DATA.in_Title_Y_Offset = INT#00) THEN
        FB_TN_SC_WRITE.Iin_Y := Xus_TN_INPUT_CONTROL_DATA.in_Y;
        FB_TN_SC_WRITE.Iin_X := Xus_TN_INPUT_CONTROL_DATA.in_X - LEN(Xus_TN_INPUT_CONTROL_DATA.st_Title_String);

      ELSE
        FB_TN_SC_WRITE.Iin_Y := Xus_TN_INPUT_CONTROL_DATA.in_Y + Xus_TN_INPUT_CONTROL_DATA.in_Title_Y_Offset;
        FB_TN_SC_WRITE.Iin_X := Xus_TN_INPUT_CONTROL_DATA.in_X + Xus_TN_INPUT_CONTROL_DATA.in_Title_X_Offset;

      END_IF;
      FB_TN_SC_WRITE.Iby_ATTR      := Xus_TN_INPUT_CONTROL_DATA.by_Title_Attr;
      FB_TN_SC_WRITE.Ist_STRING    := Xus_TN_INPUT_CONTROL_DATA.st_Title_String;
      FB_TN_SC_WRITE.Xus_TN_SCREEN := Xus_TN_SCREEN;
      FB_TN_SC_WRITE();
      Xus_TN_SCREEN := FB_TN_SC_WRITE.Xus_TN_SCREEN;

    END_IF;

    IF (Xus_TN_INPUT_CONTROL_DATA.bo_Input_Hidden = TRUE) THEN

      st_String := '';

      IF LEN(Xus_TN_INPUT_CONTROL_DATA.st_Input_Data) = LEN(Xus_TN_INPUT_CONTROL_DATA.st_Input_Mask) THEN
        FOR in_count := 1 TO LEN(Xus_TN_INPUT_CONTROL_DATA.st_Input_Data) DO

          st_CHAR := MID(Xus_TN_INPUT_CONTROL_DATA.st_Input_Mask,1,in_count);

          IF EQ_STRING(st_CHAR,' ') THEN

            st_CHAR := MID(Xus_TN_INPUT_CONTROL_DATA.st_Input_Data,1,in_count);

            IF EQ_STRING(st_CHAR,' ') THEN
              st_String := CONCAT(st_String,' ');

            ELSE
              st_String := CONCAT(st_String,'*');

            END_IF;

          ELSE
          st_CHAR := MID(Xus_TN_INPUT_CONTROL_DATA.st_Input_Data,1,in_count);
          st_String := CONCAT(st_String,st_CHAR);

          END_IF;
        END_FOR;
      END_IF;
    ELSE

      st_String := Xus_TN_INPUT_CONTROL_DATA.st_Input_Data;

    END_IF;

    IF Xus_TN_INPUT_CONTROL_DATA.bo_Focus = TRUE THEN
      by_Attr := Xus_TN_INPUT_CONTROL_DATA.by_Attr_mF;
    ELSE
      by_Attr := Xus_TN_INPUT_CONTROL_DATA.by_Attr_oF;
    END_IF;

    FB_TN_SC_WRITE.Iin_Y         := Xus_TN_INPUT_CONTROL_DATA.in_Y;
    FB_TN_SC_WRITE.Iin_X         := Xus_TN_INPUT_CONTROL_DATA.in_X;
    FB_TN_SC_WRITE.Iby_ATTR      := by_Attr;
    FB_TN_SC_WRITE.Ist_STRING    := st_String;
    FB_TN_SC_WRITE.Xus_TN_SCREEN := Xus_TN_SCREEN;
    FB_TN_SC_WRITE();
    Xus_TN_SCREEN := FB_TN_SC_WRITE.Xus_TN_SCREEN;

    Xus_TN_INPUT_CONTROL_DATA.in_Cursor_Y := Xus_TN_INPUT_CONTROL_DATA.in_Y;
    Xus_TN_INPUT_CONTROL_DATA.in_Cursor_X := Xus_TN_INPUT_CONTROL_DATA.in_X + Xus_TN_INPUT_CONTROL_DATA.in_Cursor_Pos - INT#1;

    in_old_charpos := INT#0;

    Xus_TN_INPUT_CONTROL_DATA.bo_Update_All   := FALSE;
    Xus_TN_INPUT_CONTROL_DATA.bo_Update_Input := FALSE;
  END_IF;

END_FUNCTION_BLOCK

(* ---- TN_INPUT_MENU_BAR.ST ---- *)
FUNCTION_BLOCK TN_INPUT_MENU_BAR

  VAR
    FB_TN_INPUT_MENU_POPUP :	TN_INPUT_MENU_POPUP;
    us_TN_MENU_POPUP :	us_TN_MENU_POPUP;
    FB_TN_SC_WRITE_C :	TN_SC_WRITE_C;
    ELEMENT_COUNT :	ELEMENT_COUNT;
    ELEMENT_GET :	ELEMENT_GET;
  END_VAR

  VAR
    in_ROW :	INT;
    in_COL :	INT;
    in_TITLE_Length :	INT;
    st_MENU_BAR :	oscat_STRING250;
    st_MENU_TITLE :	STRING;
    in_Count :	INT;
    in_Index :	INT;
    by_New_KeyCode :	BYTE;
    in_Scroll_Offset :	INT;
    by_ATTR :	BYTE;
    bo_Reset_Position :	BOOL;
  END_VAR

  VAR_IN_OUT
    Xus_TN_MENU :	us_TN_MENU;
    Xus_TN_SCREEN :	us_TN_SCREEN;
  END_VAR

  IF (Xus_TN_MENU.in_State = INT#00) AND (Xus_TN_MENU.bo_Create = TRUE) THEN
    Xus_TN_MENU.in_State			:= INT#01;
    Xus_TN_MENU.bo_Create			:= FALSE;
    Xus_TN_MENU.in_Menu_Selected	:= INT#00;
    Xus_TN_MENU.bo_Update			:= TRUE;
    bo_Reset_Position				:= TRUE;

    ELEMENT_GET(ELEMENT:=Xus_TN_MENU.st_MENU_TEXT,SEP:=BYTE#37,POS:=0);
    Xus_TN_MENU.st_MENU_TEXT:=ELEMENT_GET.ELEMENT;
    st_MENU_BAR:=ELEMENT_GET.ELEMENT_GET;

    ELEMENT_COUNT(SEP:=BYTE#35,ELEMENT:=st_MENU_BAR);
    st_MENU_BAR:=ELEMENT_COUNT.ELEMENT;
    Xus_TN_MENU.in_Menu_E_Count:=ELEMENT_COUNT.ELEMENT_COUNT;

  END_IF;

  by_New_KeyCode := Xus_TN_SCREEN.by_Input_Exten_Code;

  IF (by_New_KeyCode = BYTE#65) OR (by_New_KeyCode = BYTE#66) THEN
    us_TN_MENU_POPUP.by_Input_Exten_Code := by_New_KeyCode;
  ELSE
    us_TN_MENU_POPUP.by_Input_Exten_Code := BYTE#00;
  END_IF;

  IF (by_New_KeyCode = BYTE#27) THEN
    IF (Xus_TN_MENU.in_State = INT#01) AND (Xus_TN_SCREEN.bo_Modal_Dialog = FALSE) THEN
      Xus_TN_MENU.in_State := INT#02;
      Xus_TN_MENU.bo_Update := TRUE;
      Xus_TN_MENU.in_Menu_Selected := INT#00;

      Xus_TN_SCREEN.bo_Menue_Bar_Dialog := TRUE;

    ELSIF (Xus_TN_MENU.in_State = INT#02) THEN
      us_TN_MENU_POPUP.bo_Destroy	:= TRUE;
      Xus_TN_MENU.bo_Update		:= TRUE;
      Xus_TN_MENU.in_State		:= INT#01;
      bo_Reset_Position			:= TRUE;

      Xus_TN_SCREEN.bo_Menue_Bar_Dialog := FALSE;

    END_IF;
  END_IF;

  IF (Xus_TN_MENU.in_State = INT#02) THEN

    IF (by_New_KeyCode = BYTE#13)  THEN
      us_TN_MENU_POPUP.bo_Destroy	:= TRUE;
      Xus_TN_MENU.bo_Update		:= TRUE;
      Xus_TN_MENU.in_State		:= INT#01;
      bo_Reset_Position			:= TRUE;
      Xus_TN_MENU.in_Menu_Selected := (Xus_TN_MENU.in_Cur_Menu_Item * INT#10) + Xus_TN_MENU.in_Cur_Sub_Item;
      Xus_TN_SCREEN.by_Input_Exten_Code := BYTE#00;

      Xus_TN_SCREEN.bo_Menue_Bar_Dialog := FALSE;

    ELSIF (Xus_TN_MENU.bo_Destroy = TRUE) THEN
      us_TN_MENU_POPUP.bo_Destroy  := TRUE;
      Xus_TN_MENU.bo_Update        := TRUE;
      Xus_TN_MENU.in_State         := INT#01;
      bo_Reset_Position			 := TRUE;
      Xus_TN_MENU.in_Menu_Selected := INT#00;
      Xus_TN_SCREEN.by_Input_Exten_Code := BYTE#00;

      Xus_TN_SCREEN.bo_Menue_Bar_Dialog := FALSE;

    END_IF;

    IF (by_New_KeyCode = BYTE#67) THEN
      in_Scroll_Offset := INT#1;
      Xus_TN_MENU.bo_Update := TRUE;
      Xus_TN_SCREEN.by_Input_Exten_Code := BYTE#00;

    ELSIF (by_New_KeyCode = BYTE#68) THEN
      in_Scroll_Offset := INT#-1;
      Xus_TN_MENU.bo_Update := TRUE;
      Xus_TN_SCREEN.by_Input_Exten_Code := BYTE#00;
    END_IF;

  END_IF;

  IF bo_Reset_Position = TRUE THEN
    bo_Reset_Position := FALSE;
    Xus_TN_MENU.in_X_SM_old := INT#-1;
    Xus_TN_MENU.in_Y_SM_old := INT#-1;
    Xus_TN_MENU.in_X_SM_new := INT#-1;
    Xus_TN_MENU.in_Y_SM_new := INT#-1;
  END_IF;

  IF (Xus_TN_MENU.in_State > INT#00) AND (Xus_TN_MENU.bo_Update = TRUE) THEN

    Xus_TN_MENU.bo_Update := FALSE;

    in_ROW := Xus_TN_MENU.in_Y;
    in_COL := Xus_TN_MENU.in_X;

    IF in_Scroll_Offset <> INT#00 THEN
      Xus_TN_MENU.in_Cur_Menu_Item := INC2(Xus_TN_MENU.in_Cur_Menu_Item,in_Scroll_Offset,1,Xus_TN_MENU.in_Menu_E_Count);
      in_Scroll_Offset := INT#00;
    ELSE
      IF (Xus_TN_MENU.in_Cur_Menu_Item = INT#00) THEN
        Xus_TN_MENU.in_Cur_Menu_Item := INT#01;
      END_IF;
    END_IF;

    FOR in_Count := INT#01 TO Xus_TN_MENU.in_Menu_E_Count DO;

      IF (in_Count = Xus_TN_MENU.in_Cur_Menu_Item) AND (Xus_TN_MENU.in_State > INT#01 ) THEN
        by_ATTR := Xus_TN_MENU.by_Attr_mF;

        Xus_TN_MENU.in_Y_SM_new := in_ROW + INT#01;
        Xus_TN_MENU.in_X_SM_new := in_COL;

      ELSE
        by_ATTR := Xus_TN_MENU.by_Attr_oF;
      END_IF;

      ELEMENT_GET(ELEMENT:=st_MENU_BAR,SEP:=BYTE#35,POS:=in_Count-1);
    st_MENU_BAR:=ELEMENT_GET.ELEMENT;
      st_MENU_TITLE:=ELEMENT_GET.ELEMENT_GET;

      in_TITLE_Length := LEN(st_MENU_TITLE) + INT#02;

      FB_TN_SC_WRITE_C.Iin_Y         := in_ROW;
      FB_TN_SC_WRITE_C.Iin_X         := in_COL;
      FB_TN_SC_WRITE_C.Iby_ATTR      := by_ATTR;
      FB_TN_SC_WRITE_C.Iin_LENGTH    := in_TITLE_Length;
      FB_TN_SC_WRITE_C.Iin_OPTION    := INT#02;
      FB_TN_SC_WRITE_C.Ist_STRING    := st_MENU_TITLE;
      FB_TN_SC_WRITE_C.Xus_TN_SCREEN := Xus_TN_SCREEN;
      FB_TN_SC_WRITE_C();
      Xus_TN_SCREEN := FB_TN_SC_WRITE_C.Xus_TN_SCREEN;

      in_COL := in_COL + in_TITLE_Length;

    END_FOR;

  END_IF;

  IF Xus_TN_MENU.in_X_SM_new <> Xus_TN_MENU.in_X_SM_old THEN

    IF us_TN_MENU_POPUP.bo_Activ = TRUE THEN
      us_TN_MENU_POPUP.bo_Destroy := TRUE;

      FB_TN_INPUT_MENU_POPUP.Xus_TN_MENU_POPUP := us_TN_MENU_POPUP;
      FB_TN_INPUT_MENU_POPUP.Xus_TN_SCREEN     := Xus_TN_SCREEN;
      FB_TN_INPUT_MENU_POPUP();
      us_TN_MENU_POPUP := FB_TN_INPUT_MENU_POPUP.Xus_TN_MENU_POPUP;
      Xus_TN_SCREEN    := FB_TN_INPUT_MENU_POPUP.Xus_TN_SCREEN;

    END_IF;

    IF us_TN_MENU_POPUP.bo_Activ = FALSE THEN
      in_Index := Xus_TN_MENU.in_Cur_Menu_Item;

      ELEMENT_GET(ELEMENT:=Xus_TN_MENU.st_MENU_TEXT,SEP:=BYTE#37,POS:=in_Index);
    Xus_TN_MENU.st_MENU_TEXT:=ELEMENT_GET.ELEMENT;

      us_TN_MENU_POPUP.in_Y         := Xus_TN_MENU.in_Y_SM_new;
      us_TN_MENU_POPUP.in_X         := Xus_TN_MENU.in_X_SM_new;
      us_TN_MENU_POPUP.by_Attr_mF   := Xus_TN_MENU.by_Attr_mF;
      us_TN_MENU_POPUP.by_Attr_oF   := Xus_TN_MENU.by_Attr_oF;
      us_TN_MENU_POPUP.st_Menu_Text := ELEMENT_GET.ELEMENT_GET;
      us_TN_MENU_POPUP.bo_Create    := TRUE;

      Xus_TN_MENU.in_X_SM_old := Xus_TN_MENU.in_X_SM_new;
      Xus_TN_MENU.in_Y_SM_old := Xus_TN_MENU.in_Y_SM_new;

    END_IF;

  END_IF;

  FB_TN_INPUT_MENU_POPUP.Xus_TN_MENU_POPUP := us_TN_MENU_POPUP;
  FB_TN_INPUT_MENU_POPUP.Xus_TN_SCREEN     := Xus_TN_SCREEN;
  FB_TN_INPUT_MENU_POPUP();
  us_TN_MENU_POPUP := FB_TN_INPUT_MENU_POPUP.Xus_TN_MENU_POPUP;
  Xus_TN_SCREEN    := FB_TN_INPUT_MENU_POPUP.Xus_TN_SCREEN;

  Xus_TN_MENU.in_Cur_Sub_Item := us_TN_MENU_POPUP.in_Cur_Item;

  IF (Xus_TN_MENU.in_State = INT#01) THEN
    IF (Xus_TN_MENU.bo_Destroy = TRUE) THEN

      Xus_TN_MENU.in_State         := INT#00;
      Xus_TN_MENU.bo_Destroy       := FALSE;
      Xus_TN_MENU.in_Cur_Menu_Item := INT#00;
      Xus_TN_MENU.in_Cur_Sub_Item  := INT#00;

    END_IF;
  END_IF;

END_FUNCTION_BLOCK

(* ---- TN_INPUT_MENU_POPUP.ST ---- *)
FUNCTION_BLOCK TN_INPUT_MENU_POPUP

  VAR
    FB_TN_SC_AREA_SAVE :	TN_SC_AREA_SAVE;
    FB_TN_SC_AREA_RESTORE :	TN_SC_AREA_RESTORE;
    FB_TN_SC_LINE :	TN_SC_LINE;
    FB_TN_SC_ADD_SHADOW :	TN_SC_ADD_SHADOW;
    FB_TN_SC_BOX :	TN_SC_BOX;
    FB_TN_SC_WRITE_C :	TN_SC_WRITE_C;
    ELEMENT_COUNT :	ELEMENT_COUNT;
    ELEMENT_GET :	ELEMENT_GET;
  END_VAR

  VAR
    in_ROW :	INT;
    in_ROWS :	INT;
    in_COL :	INT;
    in_COLS :	INT;
    in_index :	INT;
    in_Count :	INT;
    in_Scroll_Offset :	INT;
    by_ATTR :	BYTE;
  END_VAR

  VAR_IN_OUT
    Xus_TN_MENU_POPUP :	us_TN_MENU_POPUP;
    Xus_TN_SCREEN :	us_TN_SCREEN;
  END_VAR

  IF (Xus_TN_MENU_POPUP.bo_Activ = FALSE) AND (Xus_TN_MENU_POPUP.bo_Create = TRUE) THEN
    Xus_TN_MENU_POPUP.bo_Activ         := TRUE;
    Xus_TN_MENU_POPUP.bo_Create        := FALSE;
    Xus_TN_MENU_POPUP.bo_Destroy       := FALSE;
    Xus_TN_MENU_POPUP.bo_Update        := TRUE;

    ELEMENT_COUNT(ELEMENT:=Xus_TN_MENU_POPUP.st_Menu_Text,SEP:=BYTE#35);
    Xus_TN_MENU_POPUP.st_Menu_Text:=ELEMENT_COUNT.ELEMENT;
    Xus_TN_MENU_POPUP.in_Menu_E_Count:=ELEMENT_COUNT.ELEMENT_COUNT;

    Xus_TN_MENU_POPUP.in_Rows := Xus_TN_MENU_POPUP.in_Menu_E_Count;

    Xus_TN_MENU_POPUP.in_Cols := INT#00;

    FOR in_Count := INT#01 TO Xus_TN_MENU_POPUP.in_Rows DO;

      ELEMENT_GET(ELEMENT:=Xus_TN_MENU_POPUP.st_Menu_Text,SEP:=BYTE#35,POS:=in_Count-1);
      Xus_TN_MENU_POPUP.st_Menu_Text:=ELEMENT_GET.ELEMENT;
      Xus_TN_MENU_POPUP.in_Cols:=MAX_INT(LEN(ELEMENT_GET.ELEMENT_GET),Xus_TN_MENU_POPUP.in_Cols);

    END_FOR;

    IF (Xus_TN_MENU_POPUP.in_X + Xus_TN_MENU_POPUP.in_Cols) > INT#75 THEN
      Xus_TN_MENU_POPUP.in_X := INT#79 - Xus_TN_MENU_POPUP.in_Cols - INT#04;
    END_IF;

    IF (Xus_TN_MENU_POPUP.in_Y + Xus_TN_MENU_POPUP.in_ROWS) > INT#21 THEN
      Xus_TN_MENU_POPUP.in_Y := INT#23 - Xus_TN_MENU_POPUP.in_ROWS - INT#2;
    END_IF;

    Xus_TN_SCREEN.bo_Modal_Dialog := TRUE;

    FB_TN_SC_AREA_SAVE.Iin_X1        := Xus_TN_MENU_POPUP.in_X;
    FB_TN_SC_AREA_SAVE.Iin_Y1        := Xus_TN_MENU_POPUP.in_Y;
    FB_TN_SC_AREA_SAVE.Iin_X2        := Xus_TN_MENU_POPUP.in_X + Xus_TN_MENU_POPUP.in_Cols + INT#04;
    FB_TN_SC_AREA_SAVE.Iin_Y2        := Xus_TN_MENU_POPUP.in_Y + Xus_TN_MENU_POPUP.in_Rows + INT#02;
    FB_TN_SC_AREA_SAVE.Xus_TN_SCREEN := Xus_TN_SCREEN;
    FB_TN_SC_AREA_SAVE();
    Xus_TN_SCREEN := FB_TN_SC_AREA_SAVE.Xus_TN_SCREEN;

    FB_TN_SC_BOX.Iin_X1        := Xus_TN_MENU_POPUP.in_X;
    FB_TN_SC_BOX.Iin_Y1        := Xus_TN_MENU_POPUP.in_Y;
    FB_TN_SC_BOX.Iin_X2        := Xus_TN_MENU_POPUP.in_X + Xus_TN_MENU_POPUP.in_Cols + INT#03;
    FB_TN_SC_BOX.Iin_Y2        := Xus_TN_MENU_POPUP.in_Y + Xus_TN_MENU_POPUP.in_Rows + INT#01;
    FB_TN_SC_BOX.Iby_FILL      := BYTE#32;
    FB_TN_SC_BOX.Iin_BORDER    := INT#01;
    FB_TN_SC_BOX.Iby_ATTR      := Xus_TN_MENU_POPUP.by_Attr_oF;
    FB_TN_SC_BOX.Xus_TN_SCREEN := Xus_TN_SCREEN;
    FB_TN_SC_BOX();
    Xus_TN_SCREEN := FB_TN_SC_BOX.Xus_TN_SCREEN;

    FB_TN_SC_ADD_SHADOW.Iin_X1        := Xus_TN_MENU_POPUP.in_X + INT#1;
    FB_TN_SC_ADD_SHADOW.Iin_Y1        := Xus_TN_MENU_POPUP.in_Y + INT#1;
    FB_TN_SC_ADD_SHADOW.Iin_X2        := Xus_TN_MENU_POPUP.in_X + Xus_TN_MENU_POPUP.in_Cols + INT#04;
    FB_TN_SC_ADD_SHADOW.Iin_Y2        := Xus_TN_MENU_POPUP.in_Y + Xus_TN_MENU_POPUP.in_Rows + INT#02;
    FB_TN_SC_ADD_SHADOW.Iin_OPTION    := INT#00;
    FB_TN_SC_ADD_SHADOW.Xus_TN_SCREEN := Xus_TN_SCREEN;
    FB_TN_SC_ADD_SHADOW();
    Xus_TN_SCREEN := FB_TN_SC_ADD_SHADOW.Xus_TN_SCREEN;

    in_COL  := Xus_TN_MENU_POPUP.in_X;
    in_ROW  := Xus_TN_MENU_POPUP.in_Y;
    in_ROWS := Xus_TN_MENU_POPUP.in_Rows;
    in_COLS := Xus_TN_MENU_POPUP.in_Cols;

    in_COLS := in_COLS + INT#02;

    FOR in_Count := INT#01 TO Xus_TN_MENU_POPUP.in_Menu_E_Count DO;
      in_ROW := in_ROW + INT#01;

      ELEMENT_GET(ELEMENT:=Xus_TN_MENU_POPUP.st_Menu_Text,SEP:=BYTE#35,POS:=in_Count-1);
    Xus_TN_MENU_POPUP.st_Menu_Text:=ELEMENT_GET.ELEMENT;

      IF EQ_STRING(ELEMENT_GET.ELEMENT_GET,'-') THEN

        FB_TN_SC_LINE.Iin_Y1			:= in_ROW;
        FB_TN_SC_LINE.Iin_X1			:= in_COL;
        FB_TN_SC_LINE.Iin_Y2			:= in_ROW;
        FB_TN_SC_LINE.Iin_X2			:= in_COL + in_COLS + INT#01;
        FB_TN_SC_LINE.Iby_ATTR		:= Xus_TN_MENU_POPUP.by_Attr_oF;
        FB_TN_SC_LINE.Iby_BORDER		:= BYTE#01;
        FB_TN_SC_LINE.Xus_TN_SCREEN	:= Xus_TN_SCREEN;
        FB_TN_SC_LINE();
        Xus_TN_SCREEN := FB_TN_SC_LINE.Xus_TN_SCREEN;

      END_IF;
    END_FOR;
  END_IF;

  IF (Xus_TN_MENU_POPUP.bo_Activ = TRUE) THEN

    CASE _BYTE_TO_INT(Xus_TN_MENU_POPUP.by_Input_Exten_Code) OF

    65:
      in_Scroll_Offset := INT#-1;
      Xus_TN_MENU_POPUP.bo_Update := TRUE;

    66:
      in_Scroll_Offset := INT#1;
      Xus_TN_MENU_POPUP.bo_Update := TRUE;

    13:
      Xus_TN_MENU_POPUP.bo_Destroy := TRUE;

    27:
      Xus_TN_MENU_POPUP.bo_Destroy := TRUE;
      Xus_TN_MENU_POPUP.in_Cur_Item := INT#00;

    67..68:
      Xus_TN_MENU_POPUP.bo_Destroy := TRUE;
      Xus_TN_MENU_POPUP.in_Cur_Item := INT#00;

    END_CASE;

  END_IF;

  IF (Xus_TN_MENU_POPUP.bo_Activ = TRUE) AND (Xus_TN_MENU_POPUP.bo_Update = TRUE) THEN

    Xus_TN_MENU_POPUP.bo_Update := FALSE;

    in_index := Xus_TN_MENU_POPUP.in_Cur_Item;

    IF (in_index < INT#01) OR (in_index > Xus_TN_MENU_POPUP.in_Menu_E_Count) THEN
      in_Scroll_Offset := INT#01;
      in_index := Xus_TN_MENU_POPUP.in_Menu_E_Count;
    END_IF;

    ELEMENT_GET(ELEMENT:=Xus_TN_MENU_POPUP.st_Menu_Text,SEP:=BYTE#35,POS:=in_index-1);
    Xus_TN_MENU_POPUP.st_Menu_Text:=ELEMENT_GET.ELEMENT;

    IF EQ_STRING(ELEMENT_GET.ELEMENT_GET,'-') THEN
      in_Scroll_Offset := INT#01;
    END_IF;

    IF in_Scroll_Offset <> INT#00 THEN

      FOR in_Count := INT#01 TO Xus_TN_MENU_POPUP.in_Menu_E_Count DO;

        in_index:=INC2(in_index,in_Scroll_Offset,1,Xus_TN_MENU_POPUP.in_Menu_E_Count);

        ELEMENT_GET(ELEMENT:=Xus_TN_MENU_POPUP.st_Menu_Text,SEP:=BYTE#35,POS:=in_index-1);
        Xus_TN_MENU_POPUP.st_Menu_Text:=ELEMENT_GET.ELEMENT;

        IF NE_STRING(ELEMENT_GET.ELEMENT_GET,'-') THEN
          EXIT;
        END_IF;

      END_FOR;
    END_IF;

    Xus_TN_MENU_POPUP.in_Cur_Item := in_index;
    in_Scroll_Offset := INT#00;

    in_COL  := Xus_TN_MENU_POPUP.in_X;
    in_ROW  := Xus_TN_MENU_POPUP.in_Y;
    in_ROWS := Xus_TN_MENU_POPUP.in_Rows;
    in_COLS := Xus_TN_MENU_POPUP.in_Cols;

    in_COLS := in_COLS + INT#02;

    FOR in_Count := INT#01 TO Xus_TN_MENU_POPUP.in_Menu_E_Count DO;

      in_ROW := in_ROW + INT#01;

      IF in_Count = Xus_TN_MENU_POPUP.in_Cur_Item THEN
        by_ATTR := Xus_TN_MENU_POPUP.by_Attr_mF;
      ELSE
        by_ATTR := Xus_TN_MENU_POPUP.by_Attr_oF;
      END_IF;

      ELEMENT_GET(ELEMENT:=Xus_TN_MENU_POPUP.st_Menu_Text,SEP:=BYTE#35,POS:=in_Count-1);
      Xus_TN_MENU_POPUP.st_Menu_Text:=ELEMENT_GET.ELEMENT;

      IF NE_STRING(ELEMENT_GET.ELEMENT_GET,'-') THEN

        FB_TN_SC_WRITE_C.Iin_Y         := in_ROW;
        FB_TN_SC_WRITE_C.Iin_X         := in_COL + INT#01;
        FB_TN_SC_WRITE_C.Iby_ATTR      := by_ATTR;
        FB_TN_SC_WRITE_C.Iin_LENGTH    := in_COLS;
        FB_TN_SC_WRITE_C.Iin_OPTION    := INT#02;
        FB_TN_SC_WRITE_C.Ist_STRING    := ELEMENT_GET.ELEMENT_GET;
        FB_TN_SC_WRITE_C.Xus_TN_SCREEN := Xus_TN_SCREEN;
        FB_TN_SC_WRITE_C();
        Xus_TN_SCREEN := FB_TN_SC_WRITE_C.Xus_TN_SCREEN;

      END_IF;
    END_FOR;
  END_IF;

  IF (Xus_TN_MENU_POPUP.bo_Activ = TRUE) AND (Xus_TN_MENU_POPUP.bo_Destroy = TRUE) THEN

    Xus_TN_MENU_POPUP.bo_Destroy := FALSE;
    Xus_TN_MENU_POPUP.bo_Activ   := FALSE;

    FB_TN_SC_AREA_RESTORE.Xus_TN_SCREEN := Xus_TN_SCREEN;
    FB_TN_SC_AREA_RESTORE();
    Xus_TN_SCREEN := FB_TN_SC_AREA_RESTORE.Xus_TN_SCREEN;

    Xus_TN_SCREEN.bo_Modal_Dialog := FALSE;
  END_IF;

END_FUNCTION_BLOCK

(* ---- TN_INPUT_SELECT_POPUP.ST ---- *)
FUNCTION_BLOCK TN_INPUT_SELECT_POPUP

  VAR
    in_index :	INT;
    in_Element_Count :	INT;
    by_Cur_Key :	BYTE;
    by_Attr :	BYTE;
    st_String :	STRING;
  END_VAR

  VAR
    us_TN_MENU_POPUP :	us_TN_MENU_POPUP;
    FB_TN_INPUT_MENU_POPUP :	TN_INPUT_MENU_POPUP;
    FB_TN_SC_WRITE :	TN_SC_WRITE;
    FB_FIX :	FIX;
    ELEMENT_COUNT :	ELEMENT_COUNT;
    ELEMENT_GET :	ELEMENT_GET;
  END_VAR

  VAR_IN_OUT
    Xus_TN_SCREEN :	us_TN_SCREEN;
    Xus_TN_INPUT_CONTROL_DATA :	us_TN_INPUT_CONTROL_DATA;
  END_VAR

  IF (Xus_TN_INPUT_CONTROL_DATA.bo_Focus = TRUE) THEN

    by_Cur_Key := Xus_TN_INPUT_CONTROL_DATA.by_Input_Exten_Code;

    IF (us_TN_MENU_POPUP.bo_Activ = FALSE) THEN
      us_TN_MENU_POPUP.by_Input_Exten_Code := BYTE#00;

      IF (by_Cur_Key = BYTE#13) THEN
        us_TN_MENU_POPUP.in_Y         := Xus_TN_INPUT_CONTROL_DATA.in_Y;
        us_TN_MENU_POPUP.in_X         := Xus_TN_INPUT_CONTROL_DATA.in_X;
        us_TN_MENU_POPUP.by_Attr_mF   := Xus_TN_INPUT_CONTROL_DATA.by_Attr_mF;
        us_TN_MENU_POPUP.by_Attr_oF   := Xus_TN_INPUT_CONTROL_DATA.by_Attr_oF;
        us_TN_MENU_POPUP.st_Menu_Text := Xus_TN_INPUT_CONTROL_DATA.st_Input_Data;
        us_TN_MENU_POPUP.bo_Create    := TRUE;
        us_TN_MENU_POPUP.in_Cur_Item  := INT#00;
      END_IF;

      IF (us_TN_MENU_POPUP.in_Cur_Item > INT#00) THEN
        Xus_TN_INPUT_CONTROL_DATA.in_selected      := us_TN_MENU_POPUP.in_Cur_Item;
        Xus_TN_INPUT_CONTROL_DATA.bo_Input_Entered := TRUE;
        Xus_TN_INPUT_CONTROL_DATA.bo_Update_Input  := TRUE;
        us_TN_MENU_POPUP.in_Cur_Item := INT#00;
      END_IF;

    ELSE
      us_TN_MENU_POPUP.by_Input_Exten_Code := by_Cur_Key;
    END_IF;

    FB_TN_INPUT_MENU_POPUP.Xus_TN_MENU_POPUP := us_TN_MENU_POPUP;
    FB_TN_INPUT_MENU_POPUP.Xus_TN_SCREEN     := Xus_TN_SCREEN;
    FB_TN_INPUT_MENU_POPUP();
    us_TN_MENU_POPUP := FB_TN_INPUT_MENU_POPUP.Xus_TN_MENU_POPUP;
    Xus_TN_SCREEN    := FB_TN_INPUT_MENU_POPUP.Xus_TN_SCREEN;

  END_IF;

  IF (Xus_TN_INPUT_CONTROL_DATA.bo_Update_Input = TRUE) OR (Xus_TN_INPUT_CONTROL_DATA.bo_Update_All = TRUE) THEN

    IF Xus_TN_INPUT_CONTROL_DATA.bo_Update_All = TRUE THEN

      IF (Xus_TN_INPUT_CONTROL_DATA.in_Title_X_Offset = INT#00) AND (Xus_TN_INPUT_CONTROL_DATA.in_Title_Y_Offset = INT#00) THEN
        FB_TN_SC_WRITE.Iin_Y := Xus_TN_INPUT_CONTROL_DATA.in_Y;
        FB_TN_SC_WRITE.Iin_X := Xus_TN_INPUT_CONTROL_DATA.in_X - LEN(Xus_TN_INPUT_CONTROL_DATA.st_Title_String);

      ELSE
        FB_TN_SC_WRITE.Iin_Y := Xus_TN_INPUT_CONTROL_DATA.in_Y + Xus_TN_INPUT_CONTROL_DATA.in_Title_Y_Offset;
        FB_TN_SC_WRITE.Iin_X := Xus_TN_INPUT_CONTROL_DATA.in_X + Xus_TN_INPUT_CONTROL_DATA.in_Title_X_Offset;

      END_IF;

      FB_TN_SC_WRITE.Iby_ATTR      := Xus_TN_INPUT_CONTROL_DATA.by_Title_Attr;
      FB_TN_SC_WRITE.Ist_STRING    := Xus_TN_INPUT_CONTROL_DATA.st_Title_String;
      FB_TN_SC_WRITE.Xus_TN_SCREEN := Xus_TN_SCREEN;
      FB_TN_SC_WRITE();
      Xus_TN_SCREEN := FB_TN_SC_WRITE.Xus_TN_SCREEN;

    END_IF;

    ELEMENT_COUNT(SEP:=BYTE#35,ELEMENT:=Xus_TN_INPUT_CONTROL_DATA.st_Input_Data);
    Xus_TN_INPUT_CONTROL_DATA.st_Input_Data:=ELEMENT_COUNT.ELEMENT;
    in_Element_Count:=ELEMENT_COUNT.ELEMENT_COUNT;

    IF in_Element_Count > INT#00 THEN

      Xus_TN_INPUT_CONTROL_DATA.in_selected:=LIMIT_INT(1,Xus_TN_INPUT_CONTROL_DATA.in_selected,in_Element_Count);

      in_index := Xus_TN_INPUT_CONTROL_DATA.in_selected;

      ELEMENT_GET(ELEMENT:=Xus_TN_INPUT_CONTROL_DATA.st_Input_Data,SEP:=BYTE#35,POS:=in_index-1);
      Xus_TN_INPUT_CONTROL_DATA.st_Input_Data:=ELEMENT_GET.ELEMENT;

      st_String:=ELEMENT_GET.ELEMENT_GET;

      FB_FIX.str:=st_String;
    FB_FIX.L:=LEN(Xus_TN_INPUT_CONTROL_DATA.st_Input_Mask);
    FB_FIX.C:=BYTE#32;
    FB_FIX.M:=Xus_TN_INPUT_CONTROL_DATA.in_Input_Option;
      FB_FIX();
      st_String:=FB_FIX.FIX;

      Xus_TN_INPUT_CONTROL_DATA.st_Input_String := st_String;

      IF Xus_TN_INPUT_CONTROL_DATA.bo_Focus = TRUE THEN
        by_Attr := Xus_TN_INPUT_CONTROL_DATA.by_Attr_mF;
      ELSE
        by_Attr := Xus_TN_INPUT_CONTROL_DATA.by_Attr_oF;
      END_IF;

      FB_TN_SC_WRITE.Iin_X         := Xus_TN_INPUT_CONTROL_DATA.in_X;
      FB_TN_SC_WRITE.Iin_Y         := Xus_TN_INPUT_CONTROL_DATA.in_Y;
      FB_TN_SC_WRITE.Iby_ATTR      := by_Attr;
      FB_TN_SC_WRITE.Ist_STRING    := st_String;
      FB_TN_SC_WRITE.Xus_TN_SCREEN := Xus_TN_SCREEN;
      FB_TN_SC_WRITE();
      Xus_TN_SCREEN := FB_TN_SC_WRITE.Xus_TN_SCREEN;

    END_IF;

    Xus_TN_INPUT_CONTROL_DATA.in_Cursor_X := Xus_TN_INPUT_CONTROL_DATA.in_X;
    Xus_TN_INPUT_CONTROL_DATA.in_Cursor_Y := Xus_TN_INPUT_CONTROL_DATA.in_Y;

    Xus_TN_INPUT_CONTROL_DATA.bo_Update_All   := FALSE;
    Xus_TN_INPUT_CONTROL_DATA.bo_Update_Input := FALSE;

  END_IF;

END_FUNCTION_BLOCK

(* ---- TN_INPUT_SELECT_TEXT.ST ---- *)
TYPE
  bya_TN_CHAR:       	ARRAY [0..1919] OF BYTE;
  bya_TN_BACKUP:     	ARRAY [0..1919] OF BYTE;
  bya_TN_COLOR:      	ARRAY [0..1919] OF BYTE;
  bya_TN_Line_Update:	ARRAY [0..23]   OF BOOL;

  us_TN_SCREEN :
  STRUCT
		bya_CHAR:			bya_TN_CHAR;
		bya_COLOR:			bya_TN_COLOR;
		bya_BACKUP:			bya_TN_BACKUP;
		bya_Line_Update:	bya_TN_Line_Update;

		by_Input_Exten_Code:    BYTE;
		by_Input_ASCII_Code:    BYTE;
		bo_Input_ASCII_IsNum:   BOOL;
		in_Page_Number:        	INT;
		in_Cursor_X:           	INT;
		in_Cursor_Y:           	INT;
		in_EOS_Offset:         	INT;
		by_Clear_Screen_Attr:  	BYTE;
		bo_Clear_Screen:       	BOOL;
		bo_Modal_Dialog:       	BOOL;
		bo_Menue_Bar_Dialog:   	BOOL;

  END_STRUCT;
END_TYPE

FUNCTION_BLOCK TN_INPUT_SELECT_TEXT_Block

  VAR
    in_count :	INT;
    by_Attr :	BYTE;
    st_String :	STRING;
  END_VAR

  VAR
    FB_FIX :	FIX;
    FB_TN_SC_WRITE :	TN_SC_WRITE;
    ELEMENT_COUNT :	ELEMENT_COUNT;
    ELEMENT_GET :	ELEMENT_GET;
  END_VAR

  VAR_IN_OUT
    Xus_TN_SCREEN :	us_TN_SCREEN;
    Xus_TN_INPUT_CONTROL_DATA :	us_TN_INPUT_CONTROL_DATA;
  END_VAR

  IF Xus_TN_INPUT_CONTROL_DATA.bo_Focus = TRUE THEN

    IF Xus_TN_INPUT_CONTROL_DATA.by_Input_ASCII_Code = BYTE#32 THEN
      Xus_TN_INPUT_CONTROL_DATA.in_selected := Xus_TN_INPUT_CONTROL_DATA.in_selected + INT#01;
      Xus_TN_INPUT_CONTROL_DATA.bo_Update_Input := TRUE;
    END_IF;

    IF Xus_TN_INPUT_CONTROL_DATA.by_Input_Exten_Code = BYTE#13 THEN
      Xus_TN_INPUT_CONTROL_DATA.bo_Input_Entered := TRUE;
    END_IF;

  END_IF;

  IF (Xus_TN_INPUT_CONTROL_DATA.bo_Update_Input = TRUE) OR (Xus_TN_INPUT_CONTROL_DATA.bo_Update_All = TRUE) THEN

    IF Xus_TN_INPUT_CONTROL_DATA.bo_Update_All = TRUE THEN

      IF (Xus_TN_INPUT_CONTROL_DATA.in_Title_X_Offset = INT#00) AND (Xus_TN_INPUT_CONTROL_DATA.in_Title_Y_Offset = INT#00) THEN

        FB_TN_SC_WRITE.Iin_Y := Xus_TN_INPUT_CONTROL_DATA.in_Y;
        FB_TN_SC_WRITE.Iin_X := Xus_TN_INPUT_CONTROL_DATA.in_X - LEN(Xus_TN_INPUT_CONTROL_DATA.st_Title_String);

      ELSE
        FB_TN_SC_WRITE.Iin_Y := Xus_TN_INPUT_CONTROL_DATA.in_Y + Xus_TN_INPUT_CONTROL_DATA.in_Title_Y_Offset;
        FB_TN_SC_WRITE.Iin_X := Xus_TN_INPUT_CONTROL_DATA.in_X + Xus_TN_INPUT_CONTROL_DATA.in_Title_X_Offset;

      END_IF;

      FB_TN_SC_WRITE.Iby_ATTR      := Xus_TN_INPUT_CONTROL_DATA.by_Title_Attr;
      FB_TN_SC_WRITE.Ist_STRING    := Xus_TN_INPUT_CONTROL_DATA.st_Title_String;
      FB_TN_SC_WRITE.Xus_TN_SCREEN := Xus_TN_SCREEN;
      FB_TN_SC_WRITE();
      Xus_TN_SCREEN := FB_TN_SC_WRITE.Xus_TN_SCREEN;

    END_IF;

    ELEMENT_COUNT(ELEMENT:=Xus_TN_INPUT_CONTROL_DATA.st_Input_Data,SEP:=BYTE#35);
    Xus_TN_INPUT_CONTROL_DATA.st_Input_Data:=ELEMENT_COUNT.ELEMENT;
    in_count:=ELEMENT_COUNT.ELEMENT_COUNT;

    IF in_Count > INT#00 THEN

      IF Xus_TN_INPUT_CONTROL_DATA.in_selected < INT#1 THEN
        Xus_TN_INPUT_CONTROL_DATA.in_selected := INT#01;
      END_IF;

      IF Xus_TN_INPUT_CONTROL_DATA.in_selected > in_count THEN
        Xus_TN_INPUT_CONTROL_DATA.in_selected := INT#01;
      END_IF;

      ELEMENT_GET(ELEMENT:=Xus_TN_INPUT_CONTROL_DATA.st_Input_Data,SEP:=BYTE#35,POS:=Xus_TN_INPUT_CONTROL_DATA.in_selected-1);
      Xus_TN_INPUT_CONTROL_DATA.st_Input_Data := ELEMENT_GET.ELEMENT;
      st_String:=ELEMENT_GET.ELEMENT_GET;

      FB_FIX.str:=st_String;
    FB_FIX.L:=LEN(Xus_TN_INPUT_CONTROL_DATA.st_Input_Mask);
    FB_FIX.C:=BYTE#32;
    FB_FIX.M:=Xus_TN_INPUT_CONTROL_DATA.in_Input_Option;
      FB_FIX();
      st_String:=FB_FIX.FIX;

      Xus_TN_INPUT_CONTROL_DATA.st_Input_String := st_String;

      IF Xus_TN_INPUT_CONTROL_DATA.bo_Focus = TRUE THEN
        by_Attr := Xus_TN_INPUT_CONTROL_DATA.by_Attr_mF;
      ELSE
        by_Attr := Xus_TN_INPUT_CONTROL_DATA.by_Attr_oF;
      END_IF;

      FB_TN_SC_WRITE.Iin_Y         := Xus_TN_INPUT_CONTROL_DATA.in_Y;
      FB_TN_SC_WRITE.Iin_X         := Xus_TN_INPUT_CONTROL_DATA.in_X;
      FB_TN_SC_WRITE.Iby_ATTR      := by_Attr;
      FB_TN_SC_WRITE.Ist_STRING    := st_String;
      FB_TN_SC_WRITE.Xus_TN_SCREEN := Xus_TN_SCREEN;
      FB_TN_SC_WRITE();
      Xus_TN_SCREEN := FB_TN_SC_WRITE.Xus_TN_SCREEN;

    END_IF;

    Xus_TN_INPUT_CONTROL_DATA.in_Cursor_Y := Xus_TN_INPUT_CONTROL_DATA.in_Y;
    Xus_TN_INPUT_CONTROL_DATA.in_Cursor_X := Xus_TN_INPUT_CONTROL_DATA.in_X;

    Xus_TN_INPUT_CONTROL_DATA.bo_Update_All   := FALSE;
    Xus_TN_INPUT_CONTROL_DATA.bo_Update_Input := FALSE;

  END_IF;

END_FUNCTION_BLOCK

PROGRAM program0
	VAR
		Xus_TN_SCREEN :	us_TN_SCREEN;
    Xus_TN_INPUT_CONTROL_DATA :	us_TN_INPUT_CONTROL_DATA;

		func_block : TN_INPUT_SELECT_TEXT_Block;
	END_VAR
	func_block.Xus_TN_INPUT_CONTROL_DATA := Xus_TN_INPUT_CONTROL_DATA;
	func_block.Xus_TN_SCREEN := Xus_TN_SCREEN;

	func_block();
  Xus_TN_INPUT_CONTROL_DATA  := func_block.Xus_TN_INPUT_CONTROL_DATA;
	Xus_TN_SCREEN  := func_block.Xus_TN_SCREEN;
END_PROGRAM

CONFIGURATION Config0
	RESOURCE Res0 ON PLC
		TASK task0(INTERVAL := T#20ms,PRIORITY := 0);
		PROGRAM instance0 WITH task0 : program0;
	END_RESOURCE
END_CONFIGURATION

(* ---- TN_RECEIVE.ST ---- *)
TYPE
  bya_TN_CHAR:       	ARRAY [0..1919] OF BYTE;
  bya_TN_BACKUP:     	ARRAY [0..1919] OF BYTE;
  bya_TN_COLOR:      	ARRAY [0..1919] OF BYTE;
  bya_TN_Line_Update:	ARRAY [0..23]   OF BOOL;

  us_TN_SCREEN :
  STRUCT
		bya_CHAR:			bya_TN_CHAR;
		bya_COLOR:			bya_TN_COLOR;
		bya_BACKUP:			bya_TN_BACKUP;
		bya_Line_Update:	bya_TN_Line_Update;

		by_Input_Exten_Code:    BYTE;
		by_Input_ASCII_Code:    BYTE;
		bo_Input_ASCII_IsNum:   BOOL;
		in_Page_Number:        	INT;
		in_Cursor_X:           	INT;
		in_Cursor_Y:           	INT;
		in_EOS_Offset:         	INT;
		by_Clear_Screen_Attr:  	BYTE;
		bo_Clear_Screen:       	BOOL;
		bo_Modal_Dialog:       	BOOL;
		bo_Menue_Bar_Dialog:   	BOOL;

  END_STRUCT;
END_TYPE

TYPE
  oscat_NW_BUF_LONG  : ARRAY [0..4095] OF BYTE;

  oscat_NETWORK_BUFFER :
  STRUCT
    SIZE   : UINT;
    BUFFER : oscat_NW_BUF_LONG;
  END_STRUCT;
END_TYPE

FUNCTION ISC_NUM:BOOL

	VAR_INPUT
		IN :	BYTE;
	END_VAR

	ISC_NUM := IN > BYTE#47 AND IN < BYTE#58;

END_FUNCTION

FUNCTION_BLOCK TN_RECEIVE_Block

  VAR_IN_OUT
    R_BUF :	oscat_NETWORK_BUFFER;
    Xus_TN_SCREEN :	us_TN_SCREEN;
  END_VAR

  VAR
    REQ_Size :	UINT;
    REQ1 :	BYTE;
    REQ2 :	BYTE;
    REQ3 :	BYTE;
  END_VAR

  Xus_TN_SCREEN.by_Input_ASCII_Code := BYTE#00;
  Xus_TN_SCREEN.by_Input_Exten_Code := BYTE#00;

  IF R_BUF.SIZE > UINT#0 THEN
    REQ_Size := R_BUF.SIZE;
    REQ1 := R_BUF.BUFFER[0];
    REQ2 := R_BUF.BUFFER[1];
    REQ3 := R_BUF.BUFFER[2];

    IF REQ1 = BYTE#27 AND REQ_Size >= UINT#3 THEN
      IF REQ2 = BYTE#91 THEN
        IF (REQ3 >= BYTE#65 AND REQ3 <= BYTE#68) OR (REQ3 = BYTE#72) OR (REQ3 = BYTE#75) THEN
          Xus_TN_SCREEN.by_Input_Exten_Code := REQ3;
        END_IF;
      ELSIF REQ2 = BYTE#79 THEN
        IF REQ3 >= BYTE#80 AND REQ3 <= BYTE#83 THEN
          Xus_TN_SCREEN.by_Input_Exten_Code := REQ3;
        END_IF;
      END_IF;
    ELSIF REQ1 >= BYTE#32 AND REQ1 <= BYTE#126 THEN
    Xus_TN_SCREEN.by_Input_ASCII_Code := REQ1;
      Xus_TN_SCREEN.bo_Input_ASCII_IsNum := ISC_NUM(REQ1);
    ELSIF REQ1 = BYTE#8 OR REQ1 = BYTE#9 OR REQ1 = BYTE#13 OR REQ1 = BYTE#27 THEN
    Xus_TN_SCREEN.by_Input_Exten_Code := REQ1;
    END_IF;

    R_BUF.SIZE := UINT#00;
  END_IF;

END_FUNCTION_BLOCK

PROGRAM program0
	VAR
		R_BUF :	oscat_NETWORK_BUFFER;
    Xus_TN_SCREEN :	us_TN_SCREEN;

		func_block : TN_RECEIVE_Block;
	END_VAR
	func_block.R_BUF := R_BUF;
	func_block.Xus_TN_SCREEN := Xus_TN_SCREEN;

	func_block();
  R_BUF  := func_block.R_BUF;
	Xus_TN_SCREEN  := func_block.Xus_TN_SCREEN;
END_PROGRAM

CONFIGURATION Config0
	RESOURCE Res0 ON PLC
		TASK task0(INTERVAL := T#20ms,PRIORITY := 0);
		PROGRAM instance0 WITH task0 : program0;
	END_RESOURCE
END_CONFIGURATION

(* ---- TN_SC_ADD_SHADOW.ST ---- *)
TYPE
  bya_TN_CHAR:       	ARRAY [0..1919] OF BYTE;
  bya_TN_BACKUP:     	ARRAY [0..1919] OF BYTE;
  bya_TN_COLOR:      	ARRAY [0..1919] OF BYTE;
  bya_TN_Line_Update:	ARRAY [0..23]   OF BOOL;

  us_TN_SCREEN :
  STRUCT
		bya_CHAR:			bya_TN_CHAR;
		bya_COLOR:			bya_TN_COLOR;
		bya_BACKUP:			bya_TN_BACKUP;
		bya_Line_Update:	bya_TN_Line_Update;

		by_Input_Exten_Code:    BYTE;
		by_Input_ASCII_Code:    BYTE;
		bo_Input_ASCII_IsNum:   BOOL;
		in_Page_Number:        	INT;
		in_Cursor_X:           	INT;
		in_Cursor_Y:           	INT;
		in_EOS_Offset:         	INT;
		by_Clear_Screen_Attr:  	BYTE;
		bo_Clear_Screen:       	BOOL;
		bo_Modal_Dialog:       	BOOL;
		bo_Menue_Bar_Dialog:   	BOOL;

  END_STRUCT;
END_TYPE

FUNCTION TN_SC_XY2_ERROR:BOOL

	VAR_INPUT
		X1 :	INT;
		Y1 :	INT;
		X2 :	INT;
		Y2 :	INT;
	END_VAR

	TN_SC_XY2_ERROR := Y1 < 0 OR X1 < 0 OR Y2 < 0 OR X2 < 0 OR Y1 > 23 OR X1 > 79 OR Y2 > 23 OR X2 > 79;

END_FUNCTION

FUNCTION TN_SC_SHADOW_ATTR:BYTE

	VAR_INPUT
		Iby_ATTR :	BYTE;
	END_VAR

	TN_SC_SHADOW_ATTR := ((Iby_ATTR AND BYTE#2#11110000) OR BYTE#2#00001000);

END_FUNCTION

FUNCTION_BLOCK TN_SC_ADD_SHADOW_Block

  VAR
    in_Offset :	INT;
    in_X :	INT;
    in_Y :	INT;
  END_VAR

  VAR_INPUT
    Iin_Y1 :	INT;
    Iin_X1 :	INT;
    Iin_Y2 :	INT;
    Iin_X2 :	INT;
    Iin_OPTION :	INT;
  END_VAR

  VAR_IN_OUT
    Xus_TN_SCREEN :	us_TN_SCREEN;
  END_VAR

  IF TN_SC_XY2_ERROR(Iin_X1,Iin_Y1,Iin_X2,Iin_Y2) THEN RETURN; END_IF;

  in_Offset := (Iin_Y1 * 80) + Iin_X2;

  IF Iin_OPTION = INT#00 THEN
    FOR in_Y := Iin_Y1 TO Iin_Y2 DO
      Xus_TN_SCREEN.bya_COLOR[in_Offset] := TN_SC_SHADOW_ATTR(Xus_TN_SCREEN.bya_COLOR[in_Offset]);
      in_Offset := in_Offset + 80;
      Xus_TN_SCREEN.bya_Line_Update[in_Y] := TRUE;
    END_FOR;
  ELSE
    FOR in_Y := Iin_Y1 TO Iin_Y2 DO
      Xus_TN_SCREEN.bya_COLOR[in_Offset] := BYTE#00;
      Xus_TN_SCREEN.bya_CHAR[in_Offset]  := BYTE#32;
      in_Offset := in_Offset + 80;
      Xus_TN_SCREEN.bya_Line_Update[in_Y] := TRUE;
    END_FOR;
  END_IF;

  in_Offset := (Iin_Y2 * 80) + Iin_X1;

  IF Iin_OPTION = INT#00 THEN
    FOR in_X  := Iin_X1 TO Iin_X2 DO
      Xus_TN_SCREEN.bya_COLOR[in_Offset] := TN_SC_SHADOW_ATTR(Xus_TN_SCREEN.bya_COLOR[in_Offset]);
      in_Offset := in_Offset + 1;
    END_FOR;
  ELSE
    FOR in_X  := Iin_X1 TO Iin_X2 DO
      Xus_TN_SCREEN.bya_COLOR[in_Offset] := BYTE#00;
      Xus_TN_SCREEN.bya_CHAR[in_Offset]  := BYTE#32;
      in_Offset := in_Offset + 1;
    END_FOR;
  END_IF;

END_FUNCTION_BLOCK

PROGRAM program0
	VAR
		Iin_Y1 :	INT;
    Iin_X1 :	INT;
    Iin_Y2 :	INT;
    Iin_X2 :	INT;
    Iin_OPTION :	INT;
		Xus_TN_SCREEN :	us_TN_SCREEN;

		func_block : TN_SC_ADD_SHADOW_Block;
	END_VAR
	func_block.Iin_X1 := Iin_X1;
	func_block.Iin_Y1 := Iin_Y1;
	func_block.Iin_X2 := Iin_X2;
	func_block.Iin_Y2 := Iin_Y2;
  func_block.Iin_OPTION := Iin_OPTION;
	func_block.Xus_TN_SCREEN := Xus_TN_SCREEN;

	func_block();
	Xus_TN_SCREEN  := func_block.Xus_TN_SCREEN;
END_PROGRAM

CONFIGURATION Config0
	RESOURCE Res0 ON PLC
		TASK task0(INTERVAL := T#20ms,PRIORITY := 0);
		PROGRAM instance0 WITH task0 : program0;
	END_RESOURCE
END_CONFIGURATION
